(* IEC 61131-3 sources: plc-st-coding-agent/progress/evidence/f14_v14_remaining_20261113/jobs/codex_deepseek-v4pro (part 3) *)

(* ---- public-hard-05.candidate_02.st ---- *)
(* ENGINEERING_CONTRACT
   Manual axis output: ON while its button=1, opposite command inactive, and its limit=0; OFF on release/limit (PUB001).
   Manual grip/release: ON while button=1, opposite inactive, and its limit=0; OFF on release/limit (PUB001).
   Single-step: Start edge activates next index 0..7/wraps; output held until switch; next Start advances (PUB002-PUB003).
   Single-cycle: Start edge runs 0..7; holds each output until completion; stops after left; next Start restarts (PUB004).
   Continuous: Start edge runs 0..7 and loops after left while mode selected (PUB005).
   Emergency: EmergencyStop=FALSE overrides all outputs and freezes start/progression; state is retained (PUB006).
   Index completion: 0/4 DownLimit, 1 GripLimit, 2/6 UpLimit, 3 RightLimit, 5 ReleaseLimit, 7 LeftLimit.
   Same-scan priority: E-stop highest; sequential completion advances the step before output evaluation, so the next action can start on the completed action's scan.
   Unspecified: post-E-stop resumption uses retained state; mode changes outside a mode retain sequence state.
*)
(* CONTRACT_RULES [] *)

FUNCTION_BLOCK MechanicalArmControl
VAR_INPUT
    ManualMode : BOOL;
    SingleStepMode : BOOL;
    SingleCycleMode : BOOL;
    ContinuousMode : BOOL;
    EmergencyStop : BOOL;
    Start : BOOL;
    DownButton : BOOL;
    UpButton : BOOL;
    LeftButton : BOOL;
    RightButton : BOOL;
    GripButton : BOOL;
    ReleaseButton : BOOL;
    DownLimitSwitch : BOOL;
    UpLimitSwitch : BOOL;
    LeftLimitSwitch : BOOL;
    RightLimitSwitch : BOOL;
    GripLimitSwitch : BOOL;
    ReleaseLimitSwitch : BOOL;
END_VAR
VAR_OUTPUT
    MoveDown : BOOL;
    MoveUp : BOOL;
    MoveLeft : BOOL;
    MoveRight : BOOL;
    ActivateGrip : BOOL;
    ActivateRelease : BOOL;
END_VAR
VAR
    tmp_startEdge : R_TRIG;
    tmp_autoMode : BOOL;
    tmp_autoActive : BOOL := FALSE;
    tmp_currentStep : INT := 0;
    tmp_singleNextStep : INT := 0;
    tmp_targetReached : BOOL;
    tmp_prevSelectedModeKey : INT := -1;
    tmp_selectedModeKey : INT;

    tmp_manualDownReq : BOOL;
    tmp_manualUpReq : BOOL;
    tmp_manualLeftReq : BOOL;
    tmp_manualRightReq : BOOL;
    tmp_manualGripReq : BOOL;
    tmp_manualReleaseReq : BOOL;

    tmp_autoDown : BOOL;
    tmp_autoUp : BOOL;
    tmp_autoLeft : BOOL;
    tmp_autoRight : BOOL;
    tmp_autoGrip : BOOL;
    tmp_autoRelease : BOOL;

    tmp_down : BOOL;
    tmp_up : BOOL;
    tmp_left : BOOL;
    tmp_right : BOOL;
    tmp_grip : BOOL;
    tmp_release : BOOL;
END_VAR

tmp_startEdge(CLK := Start);

tmp_manualDownReq := ManualMode AND DownButton AND NOT DownLimitSwitch;
tmp_manualUpReq := ManualMode AND UpButton AND NOT UpLimitSwitch;
tmp_manualLeftReq := ManualMode AND LeftButton AND NOT LeftLimitSwitch;
tmp_manualRightReq := ManualMode AND RightButton AND NOT RightLimitSwitch;
tmp_manualGripReq := ManualMode AND GripButton AND NOT GripLimitSwitch;
tmp_manualReleaseReq := ManualMode AND ReleaseButton AND NOT ReleaseLimitSwitch;

tmp_autoMode := SingleStepMode OR SingleCycleMode OR ContinuousMode;

tmp_selectedModeKey := 0;
IF SingleStepMode THEN
    tmp_selectedModeKey := 1;
ELSIF SingleCycleMode THEN
    tmp_selectedModeKey := 2;
ELSIF ContinuousMode THEN
    tmp_selectedModeKey := 3;
END_IF;

IF tmp_selectedModeKey <> tmp_prevSelectedModeKey THEN
    tmp_autoActive := FALSE;
    tmp_currentStep := 0;
END_IF;
tmp_prevSelectedModeKey := tmp_selectedModeKey;

IF EmergencyStop AND tmp_startEdge.Q THEN
    IF SingleStepMode THEN
        IF NOT tmp_autoActive THEN
            tmp_currentStep := tmp_singleNextStep;
            tmp_singleNextStep := (tmp_singleNextStep + 1) MOD 8;
            tmp_autoActive := TRUE;
        END_IF;
    ELSIF SingleCycleMode THEN
        IF NOT tmp_autoActive THEN
            tmp_currentStep := 0;
            tmp_autoActive := TRUE;
        END_IF;
    ELSIF ContinuousMode THEN
        IF NOT tmp_autoActive THEN
            tmp_currentStep := 0;
            tmp_autoActive := TRUE;
        END_IF;
    END_IF;
END_IF;

CASE tmp_currentStep OF
    0, 4:
        tmp_targetReached := DownLimitSwitch;
    1:
        tmp_targetReached := GripLimitSwitch;
    2, 6:
        tmp_targetReached := UpLimitSwitch;
    3:
        tmp_targetReached := RightLimitSwitch;
    5:
        tmp_targetReached := ReleaseLimitSwitch;
    7:
        tmp_targetReached := LeftLimitSwitch;
ELSE
    tmp_targetReached := FALSE;
END_CASE;

IF EmergencyStop AND tmp_autoMode AND tmp_autoActive AND tmp_targetReached THEN
    IF SingleStepMode THEN
        tmp_autoActive := FALSE;
    ELSIF SingleCycleMode THEN
        IF tmp_currentStep >= 7 THEN
            tmp_autoActive := FALSE;
            tmp_currentStep := 0;
        ELSE
            tmp_currentStep := tmp_currentStep + 1;
        END_IF;
    ELSIF ContinuousMode THEN
        IF tmp_currentStep >= 7 THEN
            tmp_currentStep := 0;
        ELSE
            tmp_currentStep := tmp_currentStep + 1;
        END_IF;
    END_IF;
END_IF;

tmp_autoDown := tmp_autoMode AND tmp_autoActive AND ((tmp_currentStep = 0) OR (tmp_currentStep = 4)) AND NOT DownLimitSwitch;
tmp_autoGrip := tmp_autoMode AND tmp_autoActive AND (tmp_currentStep = 1) AND NOT GripLimitSwitch;
tmp_autoUp := tmp_autoMode AND tmp_autoActive AND ((tmp_currentStep = 2) OR (tmp_currentStep = 6)) AND NOT UpLimitSwitch;
tmp_autoRight := tmp_autoMode AND tmp_autoActive AND (tmp_currentStep = 3) AND NOT RightLimitSwitch;
tmp_autoRelease := tmp_autoMode AND tmp_autoActive AND (tmp_currentStep = 5) AND NOT ReleaseLimitSwitch;
tmp_autoLeft := tmp_autoMode AND tmp_autoActive AND (tmp_currentStep = 7) AND NOT LeftLimitSwitch;

tmp_down := tmp_manualDownReq OR tmp_autoDown;
tmp_up := tmp_manualUpReq OR tmp_autoUp;
tmp_left := tmp_manualLeftReq OR tmp_autoLeft;
tmp_right := tmp_manualRightReq OR tmp_autoRight;
tmp_grip := tmp_manualGripReq OR tmp_autoGrip;
tmp_release := tmp_manualReleaseReq OR tmp_autoRelease;

MoveDown := tmp_down AND NOT tmp_up AND EmergencyStop;
MoveUp := tmp_up AND NOT tmp_down AND EmergencyStop;
MoveLeft := tmp_left AND NOT tmp_right AND EmergencyStop;
MoveRight := tmp_right AND NOT tmp_left AND EmergencyStop;
ActivateGrip := tmp_grip AND NOT tmp_release AND EmergencyStop;
ActivateRelease := tmp_release AND NOT tmp_grip AND EmergencyStop;

END_FUNCTION_BLOCK

(* ---- public-hard-05.patch_base_02.st ---- *)
(* ENGINEERING_CONTRACT
   Manual axis output: ON while its button=1, opposite command inactive, and its limit=0; OFF on release/limit (PUB001).
   Manual grip/release: ON while button=1, opposite inactive, and its limit=0; OFF on release/limit (PUB001).
   Single-step: Start edge activates next index 0..7/wraps; output held until switch; next Start advances (PUB002-PUB003).
   Single-cycle: Start edge runs 0..7; holds each output until completion; stops after left; next Start restarts (PUB004).
   Continuous: Start edge runs 0..7 and loops after left while mode selected (PUB005).
   Emergency: EmergencyStop=FALSE overrides all outputs and freezes start/progression; state is retained (PUB006).
   Index completion: 0/4 DownLimit, 1 GripLimit, 2/6 UpLimit, 3 RightLimit, 5 ReleaseLimit, 7 LeftLimit.
   Same-scan priority: E-stop highest; a feedback-completed action cannot energize on its completion scan; next action starts next scan.
   Unspecified: post-E-stop resumption uses retained state; mode changes outside a mode retain sequence state.
*)
(* CONTRACT_RULES [] *)

FUNCTION_BLOCK MechanicalArmControl
VAR_INPUT
    ManualMode : BOOL;
    SingleStepMode : BOOL;
    SingleCycleMode : BOOL;
    ContinuousMode : BOOL;
    EmergencyStop : BOOL;
    Start : BOOL;
    DownButton : BOOL;
    UpButton : BOOL;
    LeftButton : BOOL;
    RightButton : BOOL;
    GripButton : BOOL;
    ReleaseButton : BOOL;
    DownLimitSwitch : BOOL;
    UpLimitSwitch : BOOL;
    LeftLimitSwitch : BOOL;
    RightLimitSwitch : BOOL;
    GripLimitSwitch : BOOL;
    ReleaseLimitSwitch : BOOL;
END_VAR
VAR_OUTPUT
    MoveDown : BOOL;
    MoveUp : BOOL;
    MoveLeft : BOOL;
    MoveRight : BOOL;
    ActivateGrip : BOOL;
    ActivateRelease : BOOL;
END_VAR
VAR
    tmp_startEdge : R_TRIG;
    tmp_autoMode : BOOL;
    tmp_autoActive : BOOL := FALSE;
    tmp_currentStep : INT := 0;
    tmp_singleNextStep : INT := 0;
    tmp_targetReached : BOOL;

    tmp_manualDownReq : BOOL;
    tmp_manualUpReq : BOOL;
    tmp_manualLeftReq : BOOL;
    tmp_manualRightReq : BOOL;
    tmp_manualGripReq : BOOL;
    tmp_manualReleaseReq : BOOL;

    tmp_autoDown : BOOL;
    tmp_autoUp : BOOL;
    tmp_autoLeft : BOOL;
    tmp_autoRight : BOOL;
    tmp_autoGrip : BOOL;
    tmp_autoRelease : BOOL;

    tmp_down : BOOL;
    tmp_up : BOOL;
    tmp_left : BOOL;
    tmp_right : BOOL;
    tmp_grip : BOOL;
    tmp_release : BOOL;
END_VAR

tmp_startEdge(CLK := Start);

tmp_manualDownReq := ManualMode AND DownButton AND NOT DownLimitSwitch;
tmp_manualUpReq := ManualMode AND UpButton AND NOT UpLimitSwitch;
tmp_manualLeftReq := ManualMode AND LeftButton AND NOT LeftLimitSwitch;
tmp_manualRightReq := ManualMode AND RightButton AND NOT RightLimitSwitch;
tmp_manualGripReq := ManualMode AND GripButton AND NOT GripLimitSwitch;
tmp_manualReleaseReq := ManualMode AND ReleaseButton AND NOT ReleaseLimitSwitch;

tmp_autoMode := SingleStepMode OR SingleCycleMode OR ContinuousMode;

IF EmergencyStop AND tmp_startEdge.Q THEN
    IF SingleStepMode THEN
        IF NOT tmp_autoActive THEN
            tmp_currentStep := tmp_singleNextStep;
            tmp_singleNextStep := (tmp_singleNextStep + 1) MOD 8;
            tmp_autoActive := TRUE;
        END_IF;
    ELSIF SingleCycleMode THEN
        IF NOT tmp_autoActive THEN
            tmp_currentStep := 0;
            tmp_autoActive := TRUE;
        END_IF;
    ELSIF ContinuousMode THEN
        IF NOT tmp_autoActive THEN
            tmp_currentStep := 0;
            tmp_autoActive := TRUE;
        END_IF;
    END_IF;
END_IF;

CASE tmp_currentStep OF
    0, 4:
        tmp_targetReached := DownLimitSwitch;
    1:
        tmp_targetReached := GripLimitSwitch;
    2, 6:
        tmp_targetReached := UpLimitSwitch;
    3:
        tmp_targetReached := RightLimitSwitch;
    5:
        tmp_targetReached := ReleaseLimitSwitch;
    7:
        tmp_targetReached := LeftLimitSwitch;
ELSE
    tmp_targetReached := FALSE;
END_CASE;

tmp_autoDown := tmp_autoMode AND tmp_autoActive AND ((tmp_currentStep = 0) OR (tmp_currentStep = 4)) AND NOT DownLimitSwitch;
tmp_autoGrip := tmp_autoMode AND tmp_autoActive AND (tmp_currentStep = 1) AND NOT GripLimitSwitch;
tmp_autoUp := tmp_autoMode AND tmp_autoActive AND ((tmp_currentStep = 2) OR (tmp_currentStep = 6)) AND NOT UpLimitSwitch;
tmp_autoRight := tmp_autoMode AND tmp_autoActive AND (tmp_currentStep = 3) AND NOT RightLimitSwitch;
tmp_autoRelease := tmp_autoMode AND tmp_autoActive AND (tmp_currentStep = 5) AND NOT ReleaseLimitSwitch;
tmp_autoLeft := tmp_autoMode AND tmp_autoActive AND (tmp_currentStep = 7) AND NOT LeftLimitSwitch;

tmp_down := tmp_manualDownReq OR tmp_autoDown;
tmp_up := tmp_manualUpReq OR tmp_autoUp;
tmp_left := tmp_manualLeftReq OR tmp_autoLeft;
tmp_right := tmp_manualRightReq OR tmp_autoRight;
tmp_grip := tmp_manualGripReq OR tmp_autoGrip;
tmp_release := tmp_manualReleaseReq OR tmp_autoRelease;

MoveDown := tmp_down AND NOT tmp_up AND EmergencyStop;
MoveUp := tmp_up AND NOT tmp_down AND EmergencyStop;
MoveLeft := tmp_left AND NOT tmp_right AND EmergencyStop;
MoveRight := tmp_right AND NOT tmp_left AND EmergencyStop;
ActivateGrip := tmp_grip AND NOT tmp_release AND EmergencyStop;
ActivateRelease := tmp_release AND NOT tmp_grip AND EmergencyStop;

IF EmergencyStop AND tmp_autoMode AND tmp_autoActive AND tmp_targetReached THEN
    IF SingleStepMode THEN
        tmp_autoActive := FALSE;
    ELSIF SingleCycleMode THEN
        IF tmp_currentStep >= 7 THEN
            tmp_autoActive := FALSE;
            tmp_currentStep := 0;
        ELSE
            tmp_currentStep := tmp_currentStep + 1;
        END_IF;
    ELSIF ContinuousMode THEN
        IF tmp_currentStep >= 7 THEN
            tmp_currentStep := 0;
        ELSE
            tmp_currentStep := tmp_currentStep + 1;
        END_IF;
    END_IF;
END_IF;

END_FUNCTION_BLOCK

(* ---- public-hard-05.raw_candidate_01.st ---- *)
(* ENGINEERING_CONTRACT
   Manual axis output: ON while its button=1, opposite command inactive, and its limit=0; OFF on release/limit (PUB001).
   Manual grip/release: ON while button=1, opposite inactive, and its limit=0; OFF on release/limit (PUB001).
   Single-step: Start edge activates next index 0..7/wraps; output held until switch; next Start advances (PUB002-PUB003).
   Single-cycle: Start edge runs 0..7; holds each output until completion; stops after left; next Start restarts (PUB004).
   Continuous: Start edge runs 0..7 and loops after left while mode selected (PUB005).
   Emergency: EmergencyStop=FALSE overrides all outputs and freezes start/progression; state is retained (PUB006).
   Index completion: 0/4 DownLimit, 1 GripLimit, 2/6 UpLimit, 3 RightLimit, 5 ReleaseLimit, 7 LeftLimit.
   Same-scan priority: E-stop highest; a feedback-completed action cannot energize on its completion scan; next action starts next scan.
   Unspecified: post-E-stop resumption uses retained state; mode changes outside a mode retain sequence state.
*)
(* CONTRACT_RULES [] *)

FUNCTION_BLOCK MechanicalArmControl
VAR_INPUT
    ManualMode : BOOL;
    SingleStepMode : BOOL;
    SingleCycleMode : BOOL;
    ContinuousMode : BOOL;
    EmergencyStop : BOOL;
    Start : BOOL;
    DownButton : BOOL;
    UpButton : BOOL;
    LeftButton : BOOL;
    RightButton : BOOL;
    GripButton : BOOL;
    ReleaseButton : BOOL;
    DownLimitSwitch : BOOL;
    UpLimitSwitch : BOOL;
    LeftLimitSwitch : BOOL;
    RightLimitSwitch : BOOL;
    GripLimitSwitch : BOOL;
    ReleaseLimitSwitch : BOOL;
END_VAR
VAR_OUTPUT
    MoveDown : BOOL;
    MoveUp : BOOL;
    MoveLeft : BOOL;
    MoveRight : BOOL;
    ActivateGrip : BOOL;
    ActivateRelease : BOOL;
END_VAR
VAR
    tmp_startEdge : R_TRIG;
    tmp_autoMode : BOOL;
    tmp_autoActive : BOOL := FALSE;
    tmp_currentStep : INT := 0;
    tmp_singleNextStep : INT := 0;
    tmp_targetReached : BOOL;

    tmp_manualDownReq : BOOL;
    tmp_manualUpReq : BOOL;
    tmp_manualLeftReq : BOOL;
    tmp_manualRightReq : BOOL;
    tmp_manualGripReq : BOOL;
    tmp_manualReleaseReq : BOOL;

    tmp_autoDown : BOOL;
    tmp_autoUp : BOOL;
    tmp_autoLeft : BOOL;
    tmp_autoRight : BOOL;
    tmp_autoGrip : BOOL;
    tmp_autoRelease : BOOL;

    tmp_down : BOOL;
    tmp_up : BOOL;
    tmp_left : BOOL;
    tmp_right : BOOL;
    tmp_grip : BOOL;
    tmp_release : BOOL;
END_VAR

tmp_startEdge(CLK := Start);

tmp_manualDownReq := ManualMode AND DownButton AND NOT DownLimitSwitch;
tmp_manualUpReq := ManualMode AND UpButton AND NOT UpLimitSwitch;
tmp_manualLeftReq := ManualMode AND LeftButton AND NOT LeftLimitSwitch;
tmp_manualRightReq := ManualMode AND RightButton AND NOT RightLimitSwitch;
tmp_manualGripReq := ManualMode AND GripButton AND NOT GripLimitSwitch;
tmp_manualReleaseReq := ManualMode AND ReleaseButton AND NOT ReleaseLimitSwitch;

tmp_autoMode := SingleStepMode OR SingleCycleMode OR ContinuousMode;

IF EmergencyStop AND tmp_startEdge.Q THEN
    IF SingleStepMode THEN
        IF NOT tmp_autoActive THEN
            tmp_currentStep := tmp_singleNextStep;
            tmp_singleNextStep := (tmp_singleNextStep + 1) MOD 8;
            tmp_autoActive := TRUE;
        END_IF;
    ELSIF SingleCycleMode THEN
        IF NOT tmp_autoActive THEN
            tmp_currentStep := 0;
            tmp_autoActive := TRUE;
        END_IF;
    ELSIF ContinuousMode THEN
        IF NOT tmp_autoActive THEN
            tmp_currentStep := 0;
            tmp_autoActive := TRUE;
        END_IF;
    END_IF;
END_IF;

CASE tmp_currentStep OF
    0, 4:
        tmp_targetReached := DownLimitSwitch;
    1:
        tmp_targetReached := GripLimitSwitch;
    2, 6:
        tmp_targetReached := UpLimitSwitch;
    3:
        tmp_targetReached := RightLimitSwitch;
    5:
        tmp_targetReached := ReleaseLimitSwitch;
    7:
        tmp_targetReached := LeftLimitSwitch;
ELSE
    tmp_targetReached := FALSE;
END_CASE;

tmp_autoDown := tmp_autoMode AND tmp_autoActive AND ((tmp_currentStep = 0) OR (tmp_currentStep = 4)) AND NOT DownLimitSwitch;
tmp_autoGrip := tmp_autoMode AND tmp_autoActive AND (tmp_currentStep = 1) AND NOT GripLimitSwitch;
tmp_autoUp := tmp_autoMode AND tmp_autoActive AND ((tmp_currentStep = 2) OR (tmp_currentStep = 6)) AND NOT UpLimitSwitch;
tmp_autoRight := tmp_autoMode AND tmp_autoActive AND (tmp_currentStep = 3) AND NOT RightLimitSwitch;
tmp_autoRelease := tmp_autoMode AND tmp_autoActive AND (tmp_currentStep = 5) AND NOT ReleaseLimitSwitch;
tmp_autoLeft := tmp_autoMode AND tmp_autoActive AND (tmp_currentStep = 7) AND NOT LeftLimitSwitch;

tmp_down := tmp_manualDownReq OR tmp_autoDown;
tmp_up := tmp_manualUpReq OR tmp_autoUp;
tmp_left := tmp_manualLeftReq OR tmp_autoLeft;
tmp_right := tmp_manualRightReq OR tmp_autoRight;
tmp_grip := tmp_manualGripReq OR tmp_autoGrip;
tmp_release := tmp_manualReleaseReq OR tmp_autoRelease;

MoveDown := tmp_down AND NOT tmp_up AND EmergencyStop;
MoveUp := tmp_up AND NOT tmp_down AND EmergencyStop;
MoveLeft := tmp_left AND NOT tmp_right AND EmergencyStop;
MoveRight := tmp_right AND NOT tmp_left AND EmergencyStop;
ActivateGrip := tmp_grip AND NOT tmp_release AND EmergencyStop;
ActivateRelease := tmp_release AND NOT tmp_grip AND EmergencyStop;

IF EmergencyStop AND tmp_autoMode AND tmp_autoActive AND tmp_targetReached THEN
    IF SingleStepMode THEN
        tmp_autoActive := FALSE;
    ELSIF SingleCycleMode THEN
        IF tmp_currentStep >= 7 THEN
            tmp_autoActive := FALSE;
            tmp_currentStep := 0;
        ELSE
            tmp_currentStep := tmp_currentStep + 1;
        END_IF;
    ELSIF ContinuousMode THEN
        IF tmp_currentStep >= 7 THEN
            tmp_currentStep := 0;
        ELSE
            tmp_currentStep := tmp_currentStep + 1;
        END_IF;
    END_IF;
END_IF;

END_FUNCTION_BLOCK

(* ---- public-hard-05.raw_candidate_02.st ---- *)
(* ENGINEERING_CONTRACT
   Manual axis output: ON while its button=1, opposite command inactive, and its limit=0; OFF on release/limit (PUB001).
   Manual grip/release: ON while button=1, opposite inactive, and its limit=0; OFF on release/limit (PUB001).
   Single-step: Start edge activates next index 0..7/wraps; output held until switch; next Start advances (PUB002-PUB003).
   Single-cycle: Start edge runs 0..7; holds each output until completion; stops after left; next Start restarts (PUB004).
   Continuous: Start edge runs 0..7 and loops after left while mode selected (PUB005).
   Emergency: EmergencyStop=FALSE overrides all outputs and freezes start/progression; state is retained (PUB006).
   Index completion: 0/4 DownLimit, 1 GripLimit, 2/6 UpLimit, 3 RightLimit, 5 ReleaseLimit, 7 LeftLimit.
   Same-scan priority: E-stop highest; sequential completion advances the step before output evaluation, so the next action can start on the completed action's scan.
   Unspecified: post-E-stop resumption uses retained state; mode changes outside a mode retain sequence state.
*)
(* CONTRACT_RULES [] *)

FUNCTION_BLOCK MechanicalArmControl
VAR_INPUT
    ManualMode : BOOL;
    SingleStepMode : BOOL;
    SingleCycleMode : BOOL;
    ContinuousMode : BOOL;
    EmergencyStop : BOOL;
    Start : BOOL;
    DownButton : BOOL;
    UpButton : BOOL;
    LeftButton : BOOL;
    RightButton : BOOL;
    GripButton : BOOL;
    ReleaseButton : BOOL;
    DownLimitSwitch : BOOL;
    UpLimitSwitch : BOOL;
    LeftLimitSwitch : BOOL;
    RightLimitSwitch : BOOL;
    GripLimitSwitch : BOOL;
    ReleaseLimitSwitch : BOOL;
END_VAR
VAR_OUTPUT
    MoveDown : BOOL;
    MoveUp : BOOL;
    MoveLeft : BOOL;
    MoveRight : BOOL;
    ActivateGrip : BOOL;
    ActivateRelease : BOOL;
END_VAR
VAR
    tmp_startEdge : R_TRIG;
    tmp_autoMode : BOOL;
    tmp_autoActive : BOOL := FALSE;
    tmp_currentStep : INT := 0;
    tmp_singleNextStep : INT := 0;
    tmp_targetReached : BOOL;
    tmp_prevSelectedModeKey : INT := -1;
    tmp_selectedModeKey : INT;

    tmp_manualDownReq : BOOL;
    tmp_manualUpReq : BOOL;
    tmp_manualLeftReq : BOOL;
    tmp_manualRightReq : BOOL;
    tmp_manualGripReq : BOOL;
    tmp_manualReleaseReq : BOOL;

    tmp_autoDown : BOOL;
    tmp_autoUp : BOOL;
    tmp_autoLeft : BOOL;
    tmp_autoRight : BOOL;
    tmp_autoGrip : BOOL;
    tmp_autoRelease : BOOL;

    tmp_down : BOOL;
    tmp_up : BOOL;
    tmp_left : BOOL;
    tmp_right : BOOL;
    tmp_grip : BOOL;
    tmp_release : BOOL;
END_VAR

tmp_startEdge(CLK := Start);

tmp_manualDownReq := ManualMode AND DownButton AND NOT DownLimitSwitch;
tmp_manualUpReq := ManualMode AND UpButton AND NOT UpLimitSwitch;
tmp_manualLeftReq := ManualMode AND LeftButton AND NOT LeftLimitSwitch;
tmp_manualRightReq := ManualMode AND RightButton AND NOT RightLimitSwitch;
tmp_manualGripReq := ManualMode AND GripButton AND NOT GripLimitSwitch;
tmp_manualReleaseReq := ManualMode AND ReleaseButton AND NOT ReleaseLimitSwitch;

tmp_autoMode := SingleStepMode OR SingleCycleMode OR ContinuousMode;

tmp_selectedModeKey := 0;
IF SingleStepMode THEN
    tmp_selectedModeKey := 1;
ELSIF SingleCycleMode THEN
    tmp_selectedModeKey := 2;
ELSIF ContinuousMode THEN
    tmp_selectedModeKey := 3;
END_IF;

IF tmp_selectedModeKey <> tmp_prevSelectedModeKey THEN
    tmp_autoActive := FALSE;
    tmp_currentStep := 0;
END_IF;
tmp_prevSelectedModeKey := tmp_selectedModeKey;

IF EmergencyStop AND tmp_startEdge.Q THEN
    IF SingleStepMode THEN
        IF NOT tmp_autoActive THEN
            tmp_currentStep := tmp_singleNextStep;
            tmp_singleNextStep := (tmp_singleNextStep + 1) MOD 8;
            tmp_autoActive := TRUE;
        END_IF;
    ELSIF SingleCycleMode THEN
        IF NOT tmp_autoActive THEN
            tmp_currentStep := 0;
            tmp_autoActive := TRUE;
        END_IF;
    ELSIF ContinuousMode THEN
        IF NOT tmp_autoActive THEN
            tmp_currentStep := 0;
            tmp_autoActive := TRUE;
        END_IF;
    END_IF;
END_IF;

CASE tmp_currentStep OF
    0, 4:
        tmp_targetReached := DownLimitSwitch;
    1:
        tmp_targetReached := GripLimitSwitch;
    2, 6:
        tmp_targetReached := UpLimitSwitch;
    3:
        tmp_targetReached := RightLimitSwitch;
    5:
        tmp_targetReached := ReleaseLimitSwitch;
    7:
        tmp_targetReached := LeftLimitSwitch;
ELSE
    tmp_targetReached := FALSE;
END_CASE;

IF EmergencyStop AND tmp_autoMode AND tmp_autoActive AND tmp_targetReached THEN
    IF SingleStepMode THEN
        tmp_autoActive := FALSE;
    ELSIF SingleCycleMode THEN
        IF tmp_currentStep >= 7 THEN
            tmp_autoActive := FALSE;
            tmp_currentStep := 0;
        ELSE
            tmp_currentStep := tmp_currentStep + 1;
        END_IF;
    ELSIF ContinuousMode THEN
        IF tmp_currentStep >= 7 THEN
            tmp_currentStep := 0;
        ELSE
            tmp_currentStep := tmp_currentStep + 1;
        END_IF;
    END_IF;
END_IF;

tmp_autoDown := tmp_autoMode AND tmp_autoActive AND ((tmp_currentStep = 0) OR (tmp_currentStep = 4)) AND NOT DownLimitSwitch;
tmp_autoGrip := tmp_autoMode AND tmp_autoActive AND (tmp_currentStep = 1) AND NOT GripLimitSwitch;
tmp_autoUp := tmp_autoMode AND tmp_autoActive AND ((tmp_currentStep = 2) OR (tmp_currentStep = 6)) AND NOT UpLimitSwitch;
tmp_autoRight := tmp_autoMode AND tmp_autoActive AND (tmp_currentStep = 3) AND NOT RightLimitSwitch;
tmp_autoRelease := tmp_autoMode AND tmp_autoActive AND (tmp_currentStep = 5) AND NOT ReleaseLimitSwitch;
tmp_autoLeft := tmp_autoMode AND tmp_autoActive AND (tmp_currentStep = 7) AND NOT LeftLimitSwitch;

tmp_down := tmp_manualDownReq OR tmp_autoDown;
tmp_up := tmp_manualUpReq OR tmp_autoUp;
tmp_left := tmp_manualLeftReq OR tmp_autoLeft;
tmp_right := tmp_manualRightReq OR tmp_autoRight;
tmp_grip := tmp_manualGripReq OR tmp_autoGrip;
tmp_release := tmp_manualReleaseReq OR tmp_autoRelease;

MoveDown := tmp_down AND NOT tmp_up AND EmergencyStop;
MoveUp := tmp_up AND NOT tmp_down AND EmergencyStop;
MoveLeft := tmp_left AND NOT tmp_right AND EmergencyStop;
MoveRight := tmp_right AND NOT tmp_left AND EmergencyStop;
ActivateGrip := tmp_grip AND NOT tmp_release AND EmergencyStop;
ActivateRelease := tmp_release AND NOT tmp_grip AND EmergencyStop;

END_FUNCTION_BLOCK

(* ---- public-hard-06.candidate_01.st ---- *)
(* ENGINEERING_CONTRACT
- MotorForward/MotorReverse: manual direct from buttons, both inhibited when both are requested or Mode=1; automatic uses forward motion states only (PUB001, PUB002).
- Automatic motion: enabled by feed/cleaning/weighing/firing completion and held until the destination sensor is active; same-scan arrival has priority over completion (PUB003-PUB008).
- kick: set when weighing completes with weight<100.0 or weight>200.0; held while rejected until SensorWeight clears or Mode=0 (PUB009).
- firingTemp: updated only on a qualified weighing, REAL degrees, linear 100..200 -> 500..550; held through firing/output until unqualified, next feed, or Mode=0 (PUB009, PUB010).
- CompletionLight: active while SensorOutput in automatic output state; cleared when the product is removed or Mode=0 (PUB008).
- Weight boundary test is inclusive: qualified is 100.0 <= weight <= 200.0 (PUB009).
*)
(* CONTRACT_RULES [] *)

TYPE E_ProductionState :
(
    ST_IDLE := 0,
    ST_MOVE_TO_WASH := 1,
    ST_AT_WASH := 2,
    ST_MOVE_TO_WEIGHT := 3,
    ST_AT_WEIGHT := 4,
    ST_MOVE_TO_FIRING := 5,
    ST_AT_FIRING := 6,
    ST_MOVE_TO_OUTPUT := 7,
    ST_AT_OUTPUT := 8,
    ST_REJECTED := 9
);
END_TYPE;

FUNCTION_BLOCK ProductionControl
VAR_INPUT
    Mode : BOOL;
    ForwardButton : BOOL;
    ReverseButton : BOOL;
    SensorFeed : BOOL;
    SensorWash : BOOL;
    SensorWeight : BOOL;
    SensorFiring : BOOL;
    SensorOutput : BOOL;
    washComplete : BOOL;
    weightComplete : BOOL;
    weight : REAL;
    firingComplete : BOOL;
END_VAR
VAR_OUTPUT
    MotorForward : BOOL;
    MotorReverse : BOOL;
    kick : BOOL;
    CompletionLight : BOOL;
    firingTemp : REAL;
END_VAR
VAR
    tmp_LocalState : E_ProductionState := ST_IDLE;
    tmp_Qualified : BOOL;
    tmp_TempLatched : REAL := 0.0;
END_VAR

IF NOT Mode THEN
    MotorForward := ForwardButton AND NOT ReverseButton;
    MotorReverse := ReverseButton AND NOT ForwardButton;
    kick := FALSE;
    CompletionLight := FALSE;
    tmp_TempLatched := 0.0;
    firingTemp := 0.0;
ELSE
    MotorReverse := FALSE;

    IF tmp_LocalState = ST_IDLE THEN
        tmp_TempLatched := 0.0;
        IF SensorFeed THEN
            tmp_LocalState := ST_MOVE_TO_WASH;
        END_IF;
    ELSIF tmp_LocalState = ST_MOVE_TO_WASH THEN
        IF SensorWash THEN
            tmp_LocalState := ST_AT_WASH;
        END_IF;
    ELSIF tmp_LocalState = ST_AT_WASH THEN
        IF SensorWeight THEN
            tmp_LocalState := ST_AT_WEIGHT;
        ELSIF washComplete THEN
            tmp_LocalState := ST_MOVE_TO_WEIGHT;
        END_IF;
    ELSIF tmp_LocalState = ST_MOVE_TO_WEIGHT THEN
        IF SensorWeight THEN
            tmp_LocalState := ST_AT_WEIGHT;
        END_IF;
    ELSIF tmp_LocalState = ST_AT_WEIGHT THEN
        IF SensorFiring THEN
            tmp_LocalState := ST_AT_FIRING;
        ELSIF weightComplete THEN
            tmp_Qualified := (weight >= 100.0) AND (weight <= 200.0);
            IF tmp_Qualified THEN
                tmp_TempLatched := 500.0 + ((weight - 100.0) * 50.0) / 100.0;
                tmp_LocalState := ST_MOVE_TO_FIRING;
            ELSE
                tmp_TempLatched := 0.0;
                tmp_LocalState := ST_REJECTED;
            END_IF;
        END_IF;
    ELSIF tmp_LocalState = ST_REJECTED THEN
        IF NOT SensorWeight THEN
            tmp_TempLatched := 0.0;
            tmp_LocalState := ST_IDLE;
        END_IF;
    ELSIF tmp_LocalState = ST_MOVE_TO_FIRING THEN
        IF SensorFiring THEN
            tmp_LocalState := ST_AT_FIRING;
        END_IF;
    ELSIF tmp_LocalState = ST_AT_FIRING THEN
        IF SensorOutput THEN
            tmp_LocalState := ST_AT_OUTPUT;
        ELSIF firingComplete THEN
            tmp_LocalState := ST_MOVE_TO_OUTPUT;
        END_IF;
    ELSIF tmp_LocalState = ST_MOVE_TO_OUTPUT THEN
        IF SensorOutput THEN
            tmp_LocalState := ST_AT_OUTPUT;
        END_IF;
    ELSIF tmp_LocalState = ST_AT_OUTPUT THEN
        IF NOT SensorOutput THEN
            tmp_TempLatched := 0.0;
            tmp_LocalState := ST_IDLE;
        END_IF;
    END_IF;

    CASE tmp_LocalState OF
        ST_MOVE_TO_WASH,
        ST_MOVE_TO_WEIGHT,
        ST_MOVE_TO_FIRING,
        ST_MOVE_TO_OUTPUT:
            MotorForward := TRUE;
    ELSE
            MotorForward := FALSE;
    END_CASE;

    kick := (tmp_LocalState = ST_REJECTED);
    CompletionLight := (tmp_LocalState = ST_AT_OUTPUT) AND SensorOutput;
    firingTemp := tmp_TempLatched;
END_IF;

(* ---- public-hard-06.candidate_02.st ---- *)
(* ENGINEERING_CONTRACT
- MotorForward/MotorReverse: manual direct from buttons, both inhibited when both are requested or Mode=1; automatic uses forward motion states only (PUB001, PUB002).
- Automatic motion: enabled by feed/cleaning/weighing/firing completion and held until the destination sensor is active; same-scan arrival has priority over completion (PUB003-PUB008).
- kick: set when weighing completes with weight<100.0 or weight>200.0; held while rejected until SensorWeight clears or Mode=0 (PUB009).
- firingTemp: updated only on a qualified weighing, REAL degrees, linear 100..200 -> 500..550; held through firing/output until unqualified, next feed, or Mode=0 (PUB009, PUB010).
- CompletionLight: active while SensorOutput in automatic output state; cleared when the product is removed or Mode=0 (PUB008).
- Weight boundary test is inclusive: qualified is 100.0 <= weight <= 200.0 (PUB009).
*)
(* CONTRACT_RULES [] *)

TYPE E_ProductionState :
(
    ST_IDLE := 0,
    ST_MOVE_TO_WASH := 1,
    ST_AT_WASH := 2,
    ST_MOVE_TO_WEIGHT := 3,
    ST_AT_WEIGHT := 4,
    ST_MOVE_TO_FIRING := 5,
    ST_AT_FIRING := 6,
    ST_MOVE_TO_OUTPUT := 7,
    ST_AT_OUTPUT := 8,
    ST_REJECTED := 9
);
END_TYPE;

FUNCTION_BLOCK ProductionControl
VAR_INPUT
    Mode : BOOL;
    ForwardButton : BOOL;
    ReverseButton : BOOL;
    SensorFeed : BOOL;
    SensorWash : BOOL;
    SensorWeight : BOOL;
    SensorFiring : BOOL;
    SensorOutput : BOOL;
    washComplete : BOOL;
    weightComplete : BOOL;
    weight : REAL;
    firingComplete : BOOL;
END_VAR
VAR_OUTPUT
    MotorForward : BOOL;
    MotorReverse : BOOL;
    kick : BOOL;
    CompletionLight : BOOL;
    firingTemp : REAL;
END_VAR
VAR
    tmp_LocalState : E_ProductionState := ST_IDLE;
    tmp_Qualified : BOOL;
    tmp_TempLatched : REAL := 0.0;
END_VAR

IF NOT Mode THEN
    MotorForward := ForwardButton AND NOT ReverseButton;
    MotorReverse := ReverseButton AND NOT ForwardButton;
    kick := FALSE;
    CompletionLight := FALSE;
    tmp_TempLatched := 0.0;
    firingTemp := 0.0;
ELSE
    MotorReverse := FALSE;

    IF tmp_LocalState = ST_IDLE THEN
        tmp_TempLatched := 0.0;
        IF SensorFeed THEN
            tmp_LocalState := ST_MOVE_TO_WASH;
        END_IF;
    ELSIF tmp_LocalState = ST_MOVE_TO_WASH THEN
        IF SensorWash THEN
            tmp_LocalState := ST_AT_WASH;
        END_IF;
    ELSIF tmp_LocalState = ST_AT_WASH THEN
        IF SensorWeight THEN
            tmp_LocalState := ST_AT_WEIGHT;
        ELSIF washComplete THEN
            tmp_LocalState := ST_MOVE_TO_WEIGHT;
        END_IF;
    ELSIF tmp_LocalState = ST_MOVE_TO_WEIGHT THEN
        IF SensorWeight THEN
            tmp_LocalState := ST_AT_WEIGHT;
        END_IF;
    ELSIF tmp_LocalState = ST_AT_WEIGHT THEN
        IF SensorFiring THEN
            tmp_LocalState := ST_AT_FIRING;
        ELSIF weightComplete THEN
            tmp_Qualified := (weight >= 100.0) AND (weight <= 200.0);
            IF tmp_Qualified THEN
                tmp_TempLatched := 500.0 + ((weight - 100.0) * 50.0) / 100.0;
                tmp_LocalState := ST_MOVE_TO_FIRING;
            ELSE
                tmp_TempLatched := 0.0;
                tmp_LocalState := ST_REJECTED;
            END_IF;
        END_IF;
    ELSIF tmp_LocalState = ST_REJECTED THEN
        IF NOT SensorWeight THEN
            tmp_TempLatched := 0.0;
            tmp_LocalState := ST_IDLE;
        END_IF;
    ELSIF tmp_LocalState = ST_MOVE_TO_FIRING THEN
        IF SensorFiring THEN
            tmp_LocalState := ST_AT_FIRING;
        END_IF;
    ELSIF tmp_LocalState = ST_AT_FIRING THEN
        IF SensorOutput THEN
            tmp_LocalState := ST_AT_OUTPUT;
        ELSIF firingComplete THEN
            tmp_LocalState := ST_MOVE_TO_OUTPUT;
        END_IF;
    ELSIF tmp_LocalState = ST_MOVE_TO_OUTPUT THEN
        IF SensorOutput THEN
            tmp_LocalState := ST_AT_OUTPUT;
        END_IF;
    ELSIF tmp_LocalState = ST_AT_OUTPUT THEN
        IF NOT SensorOutput THEN
            tmp_TempLatched := 0.0;
            tmp_LocalState := ST_IDLE;
        END_IF;
    END_IF;

    CASE tmp_LocalState OF
        ST_MOVE_TO_WASH,
        ST_MOVE_TO_WEIGHT,
        ST_MOVE_TO_FIRING,
        ST_MOVE_TO_OUTPUT:
            MotorForward := TRUE;
    ELSE
            MotorForward := FALSE;
    END_CASE;

    kick := (tmp_LocalState = ST_REJECTED);
    CompletionLight := (tmp_LocalState = ST_AT_OUTPUT) AND SensorOutput;
    firingTemp := tmp_TempLatched;
END_IF;
END_FUNCTION_BLOCK

(* ---- public-hard-06.candidate_03.st ---- *)
(* ENGINEERING_CONTRACT
- MotorForward/MotorReverse: manual direct from buttons, both inhibited when both are requested or Mode=1; automatic uses forward motion states only (PUB001, PUB002).
- Automatic motion: enabled by feed/cleaning/weighing/firing completion and held until the destination sensor is active; same-scan arrival has priority over completion (PUB003-PUB008).
- kick: set when weighing completes with weight<100.0 or weight>200.0; held while rejected until SensorWeight clears or Mode=0 (PUB009).
- firingTemp: updated only on a qualified weighing, REAL degrees, linear 100..200 -> 500..550; retained until an unqualified weighing or Mode=0 (PUB009, PUB010).
- CompletionLight: active while SensorOutput in automatic output state; cleared when the product is removed or Mode=0 (PUB008).
- Weight boundary test is inclusive: qualified is 100.0 <= weight <= 200.0 (PUB009).
*)
(* CONTRACT_RULES [] *)

TYPE E_ProductionState :
(
    ST_IDLE := 0,
    ST_MOVE_TO_WASH := 1,
    ST_AT_WASH := 2,
    ST_MOVE_TO_WEIGHT := 3,
    ST_AT_WEIGHT := 4,
    ST_MOVE_TO_FIRING := 5,
    ST_AT_FIRING := 6,
    ST_MOVE_TO_OUTPUT := 7,
    ST_AT_OUTPUT := 8,
    ST_REJECTED := 9
);
END_TYPE;

FUNCTION_BLOCK ProductionControl
VAR_INPUT
    Mode : BOOL;
    ForwardButton : BOOL;
    ReverseButton : BOOL;
    SensorFeed : BOOL;
    SensorWash : BOOL;
    SensorWeight : BOOL;
    SensorFiring : BOOL;
    SensorOutput : BOOL;
    washComplete : BOOL;
    weightComplete : BOOL;
    weight : REAL;
    firingComplete : BOOL;
END_VAR
VAR_OUTPUT
    MotorForward : BOOL;
    MotorReverse : BOOL;
    kick : BOOL;
    CompletionLight : BOOL;
    firingTemp : REAL;
END_VAR
VAR
    tmp_LocalState : E_ProductionState := ST_IDLE;
    tmp_Qualified : BOOL;
    tmp_TempLatched : REAL := 0.0;
END_VAR

IF NOT Mode THEN
    MotorForward := ForwardButton AND NOT ReverseButton;
    MotorReverse := ReverseButton AND NOT ForwardButton;
    kick := FALSE;
    CompletionLight := FALSE;
    tmp_TempLatched := 0.0;
    firingTemp := 0.0;
ELSE
    MotorReverse := FALSE;

    IF tmp_LocalState = ST_IDLE THEN
        IF SensorFeed THEN
            tmp_LocalState := ST_MOVE_TO_WASH;
        END_IF;
    ELSIF tmp_LocalState = ST_MOVE_TO_WASH THEN
        IF SensorWash THEN
            tmp_LocalState := ST_AT_WASH;
        END_IF;
    ELSIF tmp_LocalState = ST_AT_WASH THEN
        IF SensorWeight THEN
            tmp_LocalState := ST_AT_WEIGHT;
        ELSIF washComplete THEN
            tmp_LocalState := ST_MOVE_TO_WEIGHT;
        END_IF;
    ELSIF tmp_LocalState = ST_MOVE_TO_WEIGHT THEN
        IF SensorWeight THEN
            tmp_LocalState := ST_AT_WEIGHT;
        END_IF;
    ELSIF tmp_LocalState = ST_AT_WEIGHT THEN
        IF SensorFiring THEN
            tmp_LocalState := ST_AT_FIRING;
        ELSIF weightComplete THEN
            tmp_Qualified := (weight >= 100.0) AND (weight <= 200.0);
            IF tmp_Qualified THEN
                tmp_TempLatched := 500.0 + ((weight - 100.0) * 50.0) / 100.0;
                tmp_LocalState := ST_MOVE_TO_FIRING;
            ELSE
                tmp_TempLatched := 0.0;
                tmp_LocalState := ST_REJECTED;
            END_IF;
        END_IF;
    ELSIF tmp_LocalState = ST_REJECTED THEN
        IF NOT SensorWeight THEN
            tmp_TempLatched := 0.0;
            tmp_LocalState := ST_IDLE;
        END_IF;
    ELSIF tmp_LocalState = ST_MOVE_TO_FIRING THEN
        IF SensorFiring THEN
            tmp_LocalState := ST_AT_FIRING;
        END_IF;
    ELSIF tmp_LocalState = ST_AT_FIRING THEN
        IF SensorOutput THEN
            tmp_LocalState := ST_AT_OUTPUT;
        ELSIF firingComplete THEN
            tmp_LocalState := ST_MOVE_TO_OUTPUT;
        END_IF;
    ELSIF tmp_LocalState = ST_MOVE_TO_OUTPUT THEN
        IF SensorOutput THEN
            tmp_LocalState := ST_AT_OUTPUT;
        END_IF;
    ELSIF tmp_LocalState = ST_AT_OUTPUT THEN
        IF NOT SensorOutput THEN
            tmp_LocalState := ST_IDLE;
        END_IF;
    END_IF;

    CASE tmp_LocalState OF
        ST_MOVE_TO_WASH,
        ST_MOVE_TO_WEIGHT,
        ST_MOVE_TO_FIRING,
        ST_MOVE_TO_OUTPUT:
            MotorForward := TRUE;
    ELSE
            MotorForward := FALSE;
    END_CASE;

    kick := (tmp_LocalState = ST_REJECTED);
    CompletionLight := (tmp_LocalState = ST_AT_OUTPUT) AND SensorOutput;
    firingTemp := tmp_TempLatched;
END_IF;
END_FUNCTION_BLOCK

(* ---- public-hard-06.candidate_04.st ---- *)
(* ENGINEERING_CONTRACT
- MotorForward/MotorReverse: manual direct from buttons, both inhibited when both are requested or Mode=1; automatic uses forward motion states only (PUB001, PUB002).
- Automatic motion: enabled by feed/cleaning/weighing/firing completion and held until the destination sensor is active; same-scan arrival has priority over completion (PUB003-PUB008).
- kick: set when weighing completes with weight<100.0 or weight>200.0; held while rejected until SensorWeight clears or Mode=0 (PUB009).
- firingTemp: updated only on a qualified weighing, REAL degrees, linear 100..200 -> 500..550; retained until Mode=0 (PUB009, PUB010).
- CompletionLight: active while SensorOutput in automatic output state; cleared when the product is removed or Mode=0 (PUB008).
- Weight boundary test is inclusive: qualified is 100.0 <= weight <= 200.0 (PUB009).
*)
(* CONTRACT_RULES [] *)

TYPE E_ProductionState :
(
    ST_IDLE := 0,
    ST_MOVE_TO_WASH := 1,
    ST_AT_WASH := 2,
    ST_MOVE_TO_WEIGHT := 3,
    ST_AT_WEIGHT := 4,
    ST_MOVE_TO_FIRING := 5,
    ST_AT_FIRING := 6,
    ST_MOVE_TO_OUTPUT := 7,
    ST_AT_OUTPUT := 8,
    ST_REJECTED := 9
);
END_TYPE;

FUNCTION_BLOCK ProductionControl
VAR_INPUT
    Mode : BOOL;
    ForwardButton : BOOL;
    ReverseButton : BOOL;
    SensorFeed : BOOL;
    SensorWash : BOOL;
    SensorWeight : BOOL;
    SensorFiring : BOOL;
    SensorOutput : BOOL;
    washComplete : BOOL;
    weightComplete : BOOL;
    weight : REAL;
    firingComplete : BOOL;
END_VAR
VAR_OUTPUT
    MotorForward : BOOL;
    MotorReverse : BOOL;
    kick : BOOL;
    CompletionLight : BOOL;
    firingTemp : REAL;
END_VAR
VAR
    tmp_LocalState : E_ProductionState := ST_IDLE;
    tmp_Qualified : BOOL;
    tmp_TempLatched : REAL := 0.0;
END_VAR

IF NOT Mode THEN
    MotorForward := ForwardButton AND NOT ReverseButton;
    MotorReverse := ReverseButton AND NOT ForwardButton;
    kick := FALSE;
    CompletionLight := FALSE;
    tmp_TempLatched := 0.0;
    firingTemp := 0.0;
ELSE
    MotorReverse := FALSE;

    IF tmp_LocalState = ST_IDLE THEN
        IF SensorFeed THEN
            tmp_LocalState := ST_MOVE_TO_WASH;
        END_IF;
    ELSIF tmp_LocalState = ST_MOVE_TO_WASH THEN
        IF SensorWash THEN
            tmp_LocalState := ST_AT_WASH;
        END_IF;
    ELSIF tmp_LocalState = ST_AT_WASH THEN
        IF SensorWeight THEN
            tmp_LocalState := ST_AT_WEIGHT;
        ELSIF washComplete THEN
            tmp_LocalState := ST_MOVE_TO_WEIGHT;
        END_IF;
    ELSIF tmp_LocalState = ST_MOVE_TO_WEIGHT THEN
        IF SensorWeight THEN
            tmp_LocalState := ST_AT_WEIGHT;
        END_IF;
    ELSIF tmp_LocalState = ST_AT_WEIGHT THEN
        IF SensorFiring THEN
            tmp_LocalState := ST_AT_FIRING;
        ELSIF weightComplete THEN
            tmp_Qualified := (weight >= 100.0) AND (weight <= 200.0);
            IF tmp_Qualified THEN
                tmp_TempLatched := 500.0 + ((weight - 100.0) * 50.0) / 100.0;
                tmp_LocalState := ST_MOVE_TO_FIRING;
            ELSE
                tmp_LocalState := ST_REJECTED;
            END_IF;
        END_IF;
    ELSIF tmp_LocalState = ST_REJECTED THEN
        IF NOT SensorWeight THEN
            tmp_TempLatched := 0.0;
            tmp_LocalState := ST_IDLE;
        END_IF;
    ELSIF tmp_LocalState = ST_MOVE_TO_FIRING THEN
        IF SensorFiring THEN
            tmp_LocalState := ST_AT_FIRING;
        END_IF;
    ELSIF tmp_LocalState = ST_AT_FIRING THEN
        IF SensorOutput THEN
            tmp_LocalState := ST_AT_OUTPUT;
        ELSIF firingComplete THEN
            tmp_LocalState := ST_MOVE_TO_OUTPUT;
        END_IF;
    ELSIF tmp_LocalState = ST_MOVE_TO_OUTPUT THEN
        IF SensorOutput THEN
            tmp_LocalState := ST_AT_OUTPUT;
        END_IF;
    ELSIF tmp_LocalState = ST_AT_OUTPUT THEN
        IF NOT SensorOutput THEN
            tmp_LocalState := ST_IDLE;
        END_IF;
    END_IF;

    CASE tmp_LocalState OF
        ST_MOVE_TO_WASH,
        ST_MOVE_TO_WEIGHT,
        ST_MOVE_TO_FIRING,
        ST_MOVE_TO_OUTPUT:
            MotorForward := TRUE;
    ELSE
            MotorForward := FALSE;
    END_CASE;

    kick := (tmp_LocalState = ST_REJECTED);
    CompletionLight := (tmp_LocalState = ST_AT_OUTPUT) AND SensorOutput;
    firingTemp := tmp_TempLatched;
END_IF;
END_FUNCTION_BLOCK

(* ---- public-hard-06.patch_base_02.st ---- *)
(* ENGINEERING_CONTRACT
- MotorForward/MotorReverse: manual direct from buttons, both inhibited when both are requested or Mode=1; automatic uses forward motion states only (PUB001, PUB002).
- Automatic motion: enabled by feed/cleaning/weighing/firing completion and held until the destination sensor is active; same-scan arrival has priority over completion (PUB003-PUB008).
- kick: set when weighing completes with weight<100.0 or weight>200.0; held while rejected until SensorWeight clears or Mode=0 (PUB009).
- firingTemp: updated only on a qualified weighing, REAL degrees, linear 100..200 -> 500..550; held through firing/output until unqualified, next feed, or Mode=0 (PUB009, PUB010).
- CompletionLight: active while SensorOutput in automatic output state; cleared when the product is removed or Mode=0 (PUB008).
- Weight boundary test is inclusive: qualified is 100.0 <= weight <= 200.0 (PUB009).
*)
(* CONTRACT_RULES [] *)

TYPE E_ProductionState :
(
    ST_IDLE := 0,
    ST_MOVE_TO_WASH := 1,
    ST_AT_WASH := 2,
    ST_MOVE_TO_WEIGHT := 3,
    ST_AT_WEIGHT := 4,
    ST_MOVE_TO_FIRING := 5,
    ST_AT_FIRING := 6,
    ST_MOVE_TO_OUTPUT := 7,
    ST_AT_OUTPUT := 8,
    ST_REJECTED := 9
);
END_TYPE;

FUNCTION_BLOCK ProductionControl
VAR_INPUT
    Mode : BOOL;
    ForwardButton : BOOL;
    ReverseButton : BOOL;
    SensorFeed : BOOL;
    SensorWash : BOOL;
    SensorWeight : BOOL;
    SensorFiring : BOOL;
    SensorOutput : BOOL;
    washComplete : BOOL;
    weightComplete : BOOL;
    weight : REAL;
    firingComplete : BOOL;
END_VAR
VAR_OUTPUT
    MotorForward : BOOL;
    MotorReverse : BOOL;
    kick : BOOL;
    CompletionLight : BOOL;
    firingTemp : REAL;
END_VAR
VAR
    tmp_LocalState : E_ProductionState := ST_IDLE;
    tmp_Qualified : BOOL;
    tmp_TempLatched : REAL := 0.0;
END_VAR

IF NOT Mode THEN
    MotorForward := ForwardButton AND NOT ReverseButton;
    MotorReverse := ReverseButton AND NOT ForwardButton;
    kick := FALSE;
    CompletionLight := FALSE;
    tmp_TempLatched := 0.0;
    firingTemp := 0.0;
ELSE
    MotorReverse := FALSE;

    IF tmp_LocalState = ST_IDLE THEN
        tmp_TempLatched := 0.0;
        IF SensorFeed THEN
            tmp_LocalState := ST_MOVE_TO_WASH;
        END_IF;
    ELSIF tmp_LocalState = ST_MOVE_TO_WASH THEN
        IF SensorWash THEN
            tmp_LocalState := ST_AT_WASH;
        END_IF;
    ELSIF tmp_LocalState = ST_AT_WASH THEN
        IF SensorWeight THEN
            tmp_LocalState := ST_AT_WEIGHT;
        ELSIF washComplete THEN
            tmp_LocalState := ST_MOVE_TO_WEIGHT;
        END_IF;
    ELSIF tmp_LocalState = ST_MOVE_TO_WEIGHT THEN
        IF SensorWeight THEN
            tmp_LocalState := ST_AT_WEIGHT;
        END_IF;
    ELSIF tmp_LocalState = ST_AT_WEIGHT THEN
        IF SensorFiring THEN
            tmp_LocalState := ST_AT_FIRING;
        ELSIF weightComplete THEN
            tmp_Qualified := (weight >= 100.0) AND (weight <= 200.0);
            IF tmp_Qualified THEN
                tmp_TempLatched := 500.0 + ((weight - 100.0) * 50.0) / 100.0;
                tmp_LocalState := ST_MOVE_TO_FIRING;
            ELSE
                tmp_TempLatched := 0.0;
                tmp_LocalState := ST_REJECTED;
            END_IF;
        END_IF;
    ELSIF tmp_LocalState = ST_REJECTED THEN
        IF NOT SensorWeight THEN
            tmp_TempLatched := 0.0;
            tmp_LocalState := ST_IDLE;
        END_IF;
    ELSIF tmp_LocalState = ST_MOVE_TO_FIRING THEN
        IF SensorFiring THEN
            tmp_LocalState := ST_AT_FIRING;
        END_IF;
    ELSIF tmp_LocalState = ST_AT_FIRING THEN
        IF SensorOutput THEN
            tmp_LocalState := ST_AT_OUTPUT;
        ELSIF firingComplete THEN
            tmp_LocalState := ST_MOVE_TO_OUTPUT;
        END_IF;
    ELSIF tmp_LocalState = ST_MOVE_TO_OUTPUT THEN
        IF SensorOutput THEN
            tmp_LocalState := ST_AT_OUTPUT;
        END_IF;
    ELSIF tmp_LocalState = ST_AT_OUTPUT THEN
        IF NOT SensorOutput THEN
            tmp_TempLatched := 0.0;
            tmp_LocalState := ST_IDLE;
        END_IF;
    END_IF;

    CASE tmp_LocalState OF
        ST_MOVE_TO_WASH,
        ST_MOVE_TO_WEIGHT,
        ST_MOVE_TO_FIRING,
        ST_MOVE_TO_OUTPUT:
            MotorForward := TRUE;
    ELSE
            MotorForward := FALSE;
    END_CASE;

    kick := (tmp_LocalState = ST_REJECTED);
    CompletionLight := (tmp_LocalState = ST_AT_OUTPUT) AND SensorOutput;
    firingTemp := tmp_TempLatched;
END_IF;

(* ---- public-hard-06.patch_base_03.st ---- *)
(* ENGINEERING_CONTRACT
- MotorForward/MotorReverse: manual direct from buttons, both inhibited when both are requested or Mode=1; automatic uses forward motion states only (PUB001, PUB002).
- Automatic motion: enabled by feed/cleaning/weighing/firing completion and held until the destination sensor is active; same-scan arrival has priority over completion (PUB003-PUB008).
- kick: set when weighing completes with weight<100.0 or weight>200.0; held while rejected until SensorWeight clears or Mode=0 (PUB009).
- firingTemp: updated only on a qualified weighing, REAL degrees, linear 100..200 -> 500..550; held through firing/output until unqualified, next feed, or Mode=0 (PUB009, PUB010).
- CompletionLight: active while SensorOutput in automatic output state; cleared when the product is removed or Mode=0 (PUB008).
- Weight boundary test is inclusive: qualified is 100.0 <= weight <= 200.0 (PUB009).
*)
(* CONTRACT_RULES [] *)

TYPE E_ProductionState :
(
    ST_IDLE := 0,
    ST_MOVE_TO_WASH := 1,
    ST_AT_WASH := 2,
    ST_MOVE_TO_WEIGHT := 3,
    ST_AT_WEIGHT := 4,
    ST_MOVE_TO_FIRING := 5,
    ST_AT_FIRING := 6,
    ST_MOVE_TO_OUTPUT := 7,
    ST_AT_OUTPUT := 8,
    ST_REJECTED := 9
);
END_TYPE;

FUNCTION_BLOCK ProductionControl
VAR_INPUT
    Mode : BOOL;
    ForwardButton : BOOL;
    ReverseButton : BOOL;
    SensorFeed : BOOL;
    SensorWash : BOOL;
    SensorWeight : BOOL;
    SensorFiring : BOOL;
    SensorOutput : BOOL;
    washComplete : BOOL;
    weightComplete : BOOL;
    weight : REAL;
    firingComplete : BOOL;
END_VAR
VAR_OUTPUT
    MotorForward : BOOL;
    MotorReverse : BOOL;
    kick : BOOL;
    CompletionLight : BOOL;
    firingTemp : REAL;
END_VAR
VAR
    tmp_LocalState : E_ProductionState := ST_IDLE;
    tmp_Qualified : BOOL;
    tmp_TempLatched : REAL := 0.0;
END_VAR

IF NOT Mode THEN
    MotorForward := ForwardButton AND NOT ReverseButton;
    MotorReverse := ReverseButton AND NOT ForwardButton;
    kick := FALSE;
    CompletionLight := FALSE;
    tmp_TempLatched := 0.0;
    firingTemp := 0.0;
ELSE
    MotorReverse := FALSE;

    IF tmp_LocalState = ST_IDLE THEN
        tmp_TempLatched := 0.0;
        IF SensorFeed THEN
            tmp_LocalState := ST_MOVE_TO_WASH;
        END_IF;
    ELSIF tmp_LocalState = ST_MOVE_TO_WASH THEN
        IF SensorWash THEN
            tmp_LocalState := ST_AT_WASH;
        END_IF;
    ELSIF tmp_LocalState = ST_AT_WASH THEN
        IF SensorWeight THEN
            tmp_LocalState := ST_AT_WEIGHT;
        ELSIF washComplete THEN
            tmp_LocalState := ST_MOVE_TO_WEIGHT;
        END_IF;
    ELSIF tmp_LocalState = ST_MOVE_TO_WEIGHT THEN
        IF SensorWeight THEN
            tmp_LocalState := ST_AT_WEIGHT;
        END_IF;
    ELSIF tmp_LocalState = ST_AT_WEIGHT THEN
        IF SensorFiring THEN
            tmp_LocalState := ST_AT_FIRING;
        ELSIF weightComplete THEN
            tmp_Qualified := (weight >= 100.0) AND (weight <= 200.0);
            IF tmp_Qualified THEN
                tmp_TempLatched := 500.0 + ((weight - 100.0) * 50.0) / 100.0;
                tmp_LocalState := ST_MOVE_TO_FIRING;
            ELSE
                tmp_TempLatched := 0.0;
                tmp_LocalState := ST_REJECTED;
            END_IF;
        END_IF;
    ELSIF tmp_LocalState = ST_REJECTED THEN
        IF NOT SensorWeight THEN
            tmp_TempLatched := 0.0;
            tmp_LocalState := ST_IDLE;
        END_IF;
    ELSIF tmp_LocalState = ST_MOVE_TO_FIRING THEN
        IF SensorFiring THEN
            tmp_LocalState := ST_AT_FIRING;
        END_IF;
    ELSIF tmp_LocalState = ST_AT_FIRING THEN
        IF SensorOutput THEN
            tmp_LocalState := ST_AT_OUTPUT;
        ELSIF firingComplete THEN
            tmp_LocalState := ST_MOVE_TO_OUTPUT;
        END_IF;
    ELSIF tmp_LocalState = ST_MOVE_TO_OUTPUT THEN
        IF SensorOutput THEN
            tmp_LocalState := ST_AT_OUTPUT;
        END_IF;
    ELSIF tmp_LocalState = ST_AT_OUTPUT THEN
        IF NOT SensorOutput THEN
            tmp_TempLatched := 0.0;
            tmp_LocalState := ST_IDLE;
        END_IF;
    END_IF;

    CASE tmp_LocalState OF
        ST_MOVE_TO_WASH,
        ST_MOVE_TO_WEIGHT,
        ST_MOVE_TO_FIRING,
        ST_MOVE_TO_OUTPUT:
            MotorForward := TRUE;
    ELSE
            MotorForward := FALSE;
    END_CASE;

    kick := (tmp_LocalState = ST_REJECTED);
    CompletionLight := (tmp_LocalState = ST_AT_OUTPUT) AND SensorOutput;
    firingTemp := tmp_TempLatched;
END_IF;
END_FUNCTION_BLOCK

(* ---- public-hard-06.patch_base_04.st ---- *)
(* ENGINEERING_CONTRACT
- MotorForward/MotorReverse: manual direct from buttons, both inhibited when both are requested or Mode=1; automatic uses forward motion states only (PUB001, PUB002).
- Automatic motion: enabled by feed/cleaning/weighing/firing completion and held until the destination sensor is active; same-scan arrival has priority over completion (PUB003-PUB008).
- kick: set when weighing completes with weight<100.0 or weight>200.0; held while rejected until SensorWeight clears or Mode=0 (PUB009).
- firingTemp: updated only on a qualified weighing, REAL degrees, linear 100..200 -> 500..550; retained until an unqualified weighing or Mode=0 (PUB009, PUB010).
- CompletionLight: active while SensorOutput in automatic output state; cleared when the product is removed or Mode=0 (PUB008).
- Weight boundary test is inclusive: qualified is 100.0 <= weight <= 200.0 (PUB009).
*)
(* CONTRACT_RULES [] *)

TYPE E_ProductionState :
(
    ST_IDLE := 0,
    ST_MOVE_TO_WASH := 1,
    ST_AT_WASH := 2,
    ST_MOVE_TO_WEIGHT := 3,
    ST_AT_WEIGHT := 4,
    ST_MOVE_TO_FIRING := 5,
    ST_AT_FIRING := 6,
    ST_MOVE_TO_OUTPUT := 7,
    ST_AT_OUTPUT := 8,
    ST_REJECTED := 9
);
END_TYPE;

FUNCTION_BLOCK ProductionControl
VAR_INPUT
    Mode : BOOL;
    ForwardButton : BOOL;
    ReverseButton : BOOL;
    SensorFeed : BOOL;
    SensorWash : BOOL;
    SensorWeight : BOOL;
    SensorFiring : BOOL;
    SensorOutput : BOOL;
    washComplete : BOOL;
    weightComplete : BOOL;
    weight : REAL;
    firingComplete : BOOL;
END_VAR
VAR_OUTPUT
    MotorForward : BOOL;
    MotorReverse : BOOL;
    kick : BOOL;
    CompletionLight : BOOL;
    firingTemp : REAL;
END_VAR
VAR
    tmp_LocalState : E_ProductionState := ST_IDLE;
    tmp_Qualified : BOOL;
    tmp_TempLatched : REAL := 0.0;
END_VAR

IF NOT Mode THEN
    MotorForward := ForwardButton AND NOT ReverseButton;
    MotorReverse := ReverseButton AND NOT ForwardButton;
    kick := FALSE;
    CompletionLight := FALSE;
    tmp_TempLatched := 0.0;
    firingTemp := 0.0;
ELSE
    MotorReverse := FALSE;

    IF tmp_LocalState = ST_IDLE THEN
        IF SensorFeed THEN
            tmp_LocalState := ST_MOVE_TO_WASH;
        END_IF;
    ELSIF tmp_LocalState = ST_MOVE_TO_WASH THEN
        IF SensorWash THEN
            tmp_LocalState := ST_AT_WASH;
        END_IF;
    ELSIF tmp_LocalState = ST_AT_WASH THEN
        IF SensorWeight THEN
            tmp_LocalState := ST_AT_WEIGHT;
        ELSIF washComplete THEN
            tmp_LocalState := ST_MOVE_TO_WEIGHT;
        END_IF;
    ELSIF tmp_LocalState = ST_MOVE_TO_WEIGHT THEN
        IF SensorWeight THEN
            tmp_LocalState := ST_AT_WEIGHT;
        END_IF;
    ELSIF tmp_LocalState = ST_AT_WEIGHT THEN
        IF SensorFiring THEN
            tmp_LocalState := ST_AT_FIRING;
        ELSIF weightComplete THEN
            tmp_Qualified := (weight >= 100.0) AND (weight <= 200.0);
            IF tmp_Qualified THEN
                tmp_TempLatched := 500.0 + ((weight - 100.0) * 50.0) / 100.0;
                tmp_LocalState := ST_MOVE_TO_FIRING;
            ELSE
                tmp_TempLatched := 0.0;
                tmp_LocalState := ST_REJECTED;
            END_IF;
        END_IF;
    ELSIF tmp_LocalState = ST_REJECTED THEN
        IF NOT SensorWeight THEN
            tmp_TempLatched := 0.0;
            tmp_LocalState := ST_IDLE;
        END_IF;
    ELSIF tmp_LocalState = ST_MOVE_TO_FIRING THEN
        IF SensorFiring THEN
            tmp_LocalState := ST_AT_FIRING;
        END_IF;
    ELSIF tmp_LocalState = ST_AT_FIRING THEN
        IF SensorOutput THEN
            tmp_LocalState := ST_AT_OUTPUT;
        ELSIF firingComplete THEN
            tmp_LocalState := ST_MOVE_TO_OUTPUT;
        END_IF;
    ELSIF tmp_LocalState = ST_MOVE_TO_OUTPUT THEN
        IF SensorOutput THEN
            tmp_LocalState := ST_AT_OUTPUT;
        END_IF;
    ELSIF tmp_LocalState = ST_AT_OUTPUT THEN
        IF NOT SensorOutput THEN
            tmp_LocalState := ST_IDLE;
        END_IF;
    END_IF;

    CASE tmp_LocalState OF
        ST_MOVE_TO_WASH,
        ST_MOVE_TO_WEIGHT,
        ST_MOVE_TO_FIRING,
        ST_MOVE_TO_OUTPUT:
            MotorForward := TRUE;
    ELSE
            MotorForward := FALSE;
    END_CASE;

    kick := (tmp_LocalState = ST_REJECTED);
    CompletionLight := (tmp_LocalState = ST_AT_OUTPUT) AND SensorOutput;
    firingTemp := tmp_TempLatched;
END_IF;
END_FUNCTION_BLOCK

(* ---- public-hard-06.raw_candidate_01.st ---- *)
(* ENGINEERING_CONTRACT
- MotorForward/MotorReverse: manual direct from buttons, both inhibited when both are requested or Mode=1; automatic uses forward motion states only (PUB001, PUB002).
- Automatic motion: enabled by feed/cleaning/weighing/firing completion and held until the destination sensor is active; same-scan arrival has priority over completion (PUB003-PUB008).
- kick: set when weighing completes with weight<100.0 or weight>200.0; held while rejected until SensorWeight clears or Mode=0 (PUB009).
- firingTemp: updated only on a qualified weighing, REAL degrees, linear 100..200 -> 500..550; held through firing/output until unqualified, next feed, or Mode=0 (PUB009, PUB010).
- CompletionLight: active while SensorOutput in automatic output state; cleared when the product is removed or Mode=0 (PUB008).
- Weight boundary test is inclusive: qualified is 100.0 <= weight <= 200.0 (PUB009).
*)
(* CONTRACT_RULES [] *)

TYPE E_ProductionState :
(
    ST_IDLE := 0,
    ST_MOVE_TO_WASH := 1,
    ST_AT_WASH := 2,
    ST_MOVE_TO_WEIGHT := 3,
    ST_AT_WEIGHT := 4,
    ST_MOVE_TO_FIRING := 5,
    ST_AT_FIRING := 6,
    ST_MOVE_TO_OUTPUT := 7,
    ST_AT_OUTPUT := 8,
    ST_REJECTED := 9
);
END_TYPE

FUNCTION_BLOCK ProductionControl
VAR_INPUT
    Mode : BOOL;
    ForwardButton : BOOL;
    ReverseButton : BOOL;
    SensorFeed : BOOL;
    SensorWash : BOOL;
    SensorWeight : BOOL;
    SensorFiring : BOOL;
    SensorOutput : BOOL;
    washComplete : BOOL;
    weightComplete : BOOL;
    weight : REAL;
    firingComplete : BOOL;
END_VAR
VAR_OUTPUT
    MotorForward : BOOL;
    MotorReverse : BOOL;
    kick : BOOL;
    CompletionLight : BOOL;
    firingTemp : REAL;
END_VAR
VAR
    tmp_LocalState : E_ProductionState := ST_IDLE;
    tmp_Qualified : BOOL;
    tmp_TempLatched : REAL := 0.0;
END_VAR

IF NOT Mode THEN
    MotorForward := ForwardButton AND NOT ReverseButton;
    MotorReverse := ReverseButton AND NOT ForwardButton;
    kick := FALSE;
    CompletionLight := FALSE;
    tmp_TempLatched := 0.0;
    firingTemp := 0.0;
ELSE
    MotorReverse := FALSE;

    IF tmp_LocalState = ST_IDLE THEN
        tmp_TempLatched := 0.0;
        IF SensorFeed THEN
            tmp_LocalState := ST_MOVE_TO_WASH;
        END_IF;
    ELSIF tmp_LocalState = ST_MOVE_TO_WASH THEN
        IF SensorWash THEN
            tmp_LocalState := ST_AT_WASH;
        END_IF;
    ELSIF tmp_LocalState = ST_AT_WASH THEN
        IF SensorWeight THEN
            tmp_LocalState := ST_AT_WEIGHT;
        ELSIF washComplete THEN
            tmp_LocalState := ST_MOVE_TO_WEIGHT;
        END_IF;
    ELSIF tmp_LocalState = ST_MOVE_TO_WEIGHT THEN
        IF SensorWeight THEN
            tmp_LocalState := ST_AT_WEIGHT;
        END_IF;
    ELSIF tmp_LocalState = ST_AT_WEIGHT THEN
        IF SensorFiring THEN
            tmp_LocalState := ST_AT_FIRING;
        ELSIF weightComplete THEN
            tmp_Qualified := (weight >= 100.0) AND (weight <= 200.0);
            IF tmp_Qualified THEN
                tmp_TempLatched := 500.0 + ((weight - 100.0) * 50.0) / 100.0;
                tmp_LocalState := ST_MOVE_TO_FIRING;
            ELSE
                tmp_TempLatched := 0.0;
                tmp_LocalState := ST_REJECTED;
            END_IF;
        END_IF;
    ELSIF tmp_LocalState = ST_REJECTED THEN
        IF NOT SensorWeight THEN
            tmp_TempLatched := 0.0;
            tmp_LocalState := ST_IDLE;
        END_IF;
    ELSIF tmp_LocalState = ST_MOVE_TO_FIRING THEN
        IF SensorFiring THEN
            tmp_LocalState := ST_AT_FIRING;
        END_IF;
    ELSIF tmp_LocalState = ST_AT_FIRING THEN
        IF SensorOutput THEN
            tmp_LocalState := ST_AT_OUTPUT;
        ELSIF firingComplete THEN
            tmp_LocalState := ST_MOVE_TO_OUTPUT;
        END_IF;
    ELSIF tmp_LocalState = ST_MOVE_TO_OUTPUT THEN
        IF SensorOutput THEN
            tmp_LocalState := ST_AT_OUTPUT;
        END_IF;
    ELSIF tmp_LocalState = ST_AT_OUTPUT THEN
        IF NOT SensorOutput THEN
            tmp_TempLatched := 0.0;
            tmp_LocalState := ST_IDLE;
        END_IF;
    END_IF;

    CASE tmp_LocalState OF
        ST_MOVE_TO_WASH,
        ST_MOVE_TO_WEIGHT,
        ST_MOVE_TO_FIRING,
        ST_MOVE_TO_OUTPUT:
            MotorForward := TRUE;
    ELSE
            MotorForward := FALSE;
    END_CASE;

    kick := (tmp_LocalState = ST_REJECTED);
    CompletionLight := (tmp_LocalState = ST_AT_OUTPUT) AND SensorOutput;
    firingTemp := tmp_TempLatched;
END_IF;

(* ---- public-hard-06.raw_candidate_02.st ---- *)
(* ENGINEERING_CONTRACT
- MotorForward/MotorReverse: manual direct from buttons, both inhibited when both are requested or Mode=1; automatic uses forward motion states only (PUB001, PUB002).
- Automatic motion: enabled by feed/cleaning/weighing/firing completion and held until the destination sensor is active; same-scan arrival has priority over completion (PUB003-PUB008).
- kick: set when weighing completes with weight<100.0 or weight>200.0; held while rejected until SensorWeight clears or Mode=0 (PUB009).
- firingTemp: updated only on a qualified weighing, REAL degrees, linear 100..200 -> 500..550; held through firing/output until unqualified, next feed, or Mode=0 (PUB009, PUB010).
- CompletionLight: active while SensorOutput in automatic output state; cleared when the product is removed or Mode=0 (PUB008).
- Weight boundary test is inclusive: qualified is 100.0 <= weight <= 200.0 (PUB009).
*)
(* CONTRACT_RULES [] *)

TYPE E_ProductionState :
(
    ST_IDLE := 0,
    ST_MOVE_TO_WASH := 1,
    ST_AT_WASH := 2,
    ST_MOVE_TO_WEIGHT := 3,
    ST_AT_WEIGHT := 4,
    ST_MOVE_TO_FIRING := 5,
    ST_AT_FIRING := 6,
    ST_MOVE_TO_OUTPUT := 7,
    ST_AT_OUTPUT := 8,
    ST_REJECTED := 9
);
END_TYPE;

FUNCTION_BLOCK ProductionControl
VAR_INPUT
    Mode : BOOL;
    ForwardButton : BOOL;
    ReverseButton : BOOL;
    SensorFeed : BOOL;
    SensorWash : BOOL;
    SensorWeight : BOOL;
    SensorFiring : BOOL;
    SensorOutput : BOOL;
    washComplete : BOOL;
    weightComplete : BOOL;
    weight : REAL;
    firingComplete : BOOL;
END_VAR
VAR_OUTPUT
    MotorForward : BOOL;
    MotorReverse : BOOL;
    kick : BOOL;
    CompletionLight : BOOL;
    firingTemp : REAL;
END_VAR
VAR
    tmp_LocalState : E_ProductionState := ST_IDLE;
    tmp_Qualified : BOOL;
    tmp_TempLatched : REAL := 0.0;
END_VAR

IF NOT Mode THEN
    MotorForward := ForwardButton AND NOT ReverseButton;
    MotorReverse := ReverseButton AND NOT ForwardButton;
    kick := FALSE;
    CompletionLight := FALSE;
    tmp_TempLatched := 0.0;
    firingTemp := 0.0;
ELSE
    MotorReverse := FALSE;

    IF tmp_LocalState = ST_IDLE THEN
        tmp_TempLatched := 0.0;
        IF SensorFeed THEN
            tmp_LocalState := ST_MOVE_TO_WASH;
        END_IF;
    ELSIF tmp_LocalState = ST_MOVE_TO_WASH THEN
        IF SensorWash THEN
            tmp_LocalState := ST_AT_WASH;
        END_IF;
    ELSIF tmp_LocalState = ST_AT_WASH THEN
        IF SensorWeight THEN
            tmp_LocalState := ST_AT_WEIGHT;
        ELSIF washComplete THEN
            tmp_LocalState := ST_MOVE_TO_WEIGHT;
        END_IF;
    ELSIF tmp_LocalState = ST_MOVE_TO_WEIGHT THEN
        IF SensorWeight THEN
            tmp_LocalState := ST_AT_WEIGHT;
        END_IF;
    ELSIF tmp_LocalState = ST_AT_WEIGHT THEN
        IF SensorFiring THEN
            tmp_LocalState := ST_AT_FIRING;
        ELSIF weightComplete THEN
            tmp_Qualified := (weight >= 100.0) AND (weight <= 200.0);
            IF tmp_Qualified THEN
                tmp_TempLatched := 500.0 + ((weight - 100.0) * 50.0) / 100.0;
                tmp_LocalState := ST_MOVE_TO_FIRING;
            ELSE
                tmp_TempLatched := 0.0;
                tmp_LocalState := ST_REJECTED;
            END_IF;
        END_IF;
    ELSIF tmp_LocalState = ST_REJECTED THEN
        IF NOT SensorWeight THEN
            tmp_TempLatched := 0.0;
            tmp_LocalState := ST_IDLE;
        END_IF;
    ELSIF tmp_LocalState = ST_MOVE_TO_FIRING THEN
        IF SensorFiring THEN
            tmp_LocalState := ST_AT_FIRING;
        END_IF;
    ELSIF tmp_LocalState = ST_AT_FIRING THEN
        IF SensorOutput THEN
            tmp_LocalState := ST_AT_OUTPUT;
        ELSIF firingComplete THEN
            tmp_LocalState := ST_MOVE_TO_OUTPUT;
        END_IF;
    ELSIF tmp_LocalState = ST_MOVE_TO_OUTPUT THEN
        IF SensorOutput THEN
            tmp_LocalState := ST_AT_OUTPUT;
        END_IF;
    ELSIF tmp_LocalState = ST_AT_OUTPUT THEN
        IF NOT SensorOutput THEN
            tmp_TempLatched := 0.0;
            tmp_LocalState := ST_IDLE;
        END_IF;
    END_IF;

    CASE tmp_LocalState OF
        ST_MOVE_TO_WASH,
        ST_MOVE_TO_WEIGHT,
        ST_MOVE_TO_FIRING,
        ST_MOVE_TO_OUTPUT:
            MotorForward := TRUE;
    ELSE
            MotorForward := FALSE;
    END_CASE;

    kick := (tmp_LocalState = ST_REJECTED);
    CompletionLight := (tmp_LocalState = ST_AT_OUTPUT) AND SensorOutput;
    firingTemp := tmp_TempLatched;
END_IF;
END_FUNCTION_BLOCK

(* ---- public-hard-06.raw_candidate_03.st ---- *)
(* ENGINEERING_CONTRACT
- MotorForward/MotorReverse: manual direct from buttons, both inhibited when both are requested or Mode=1; automatic uses forward motion states only (PUB001, PUB002).
- Automatic motion: enabled by feed/cleaning/weighing/firing completion and held until the destination sensor is active; same-scan arrival has priority over completion (PUB003-PUB008).
- kick: set when weighing completes with weight<100.0 or weight>200.0; held while rejected until SensorWeight clears or Mode=0 (PUB009).
- firingTemp: updated only on a qualified weighing, REAL degrees, linear 100..200 -> 500..550; retained until an unqualified weighing or Mode=0 (PUB009, PUB010).
- CompletionLight: active while SensorOutput in automatic output state; cleared when the product is removed or Mode=0 (PUB008).
- Weight boundary test is inclusive: qualified is 100.0 <= weight <= 200.0 (PUB009).
*)
(* CONTRACT_RULES [] *)

TYPE E_ProductionState :
(
    ST_IDLE := 0,
    ST_MOVE_TO_WASH := 1,
    ST_AT_WASH := 2,
    ST_MOVE_TO_WEIGHT := 3,
    ST_AT_WEIGHT := 4,
    ST_MOVE_TO_FIRING := 5,
    ST_AT_FIRING := 6,
    ST_MOVE_TO_OUTPUT := 7,
    ST_AT_OUTPUT := 8,
    ST_REJECTED := 9
);
END_TYPE;

FUNCTION_BLOCK ProductionControl
VAR_INPUT
    Mode : BOOL;
    ForwardButton : BOOL;
    ReverseButton : BOOL;
    SensorFeed : BOOL;
    SensorWash : BOOL;
    SensorWeight : BOOL;
    SensorFiring : BOOL;
    SensorOutput : BOOL;
    washComplete : BOOL;
    weightComplete : BOOL;
    weight : REAL;
    firingComplete : BOOL;
END_VAR
VAR_OUTPUT
    MotorForward : BOOL;
    MotorReverse : BOOL;
    kick : BOOL;
    CompletionLight : BOOL;
    firingTemp : REAL;
END_VAR
VAR
    tmp_LocalState : E_ProductionState := ST_IDLE;
    tmp_Qualified : BOOL;
    tmp_TempLatched : REAL := 0.0;
END_VAR

IF NOT Mode THEN
    MotorForward := ForwardButton AND NOT ReverseButton;
    MotorReverse := ReverseButton AND NOT ForwardButton;
    kick := FALSE;
    CompletionLight := FALSE;
    tmp_TempLatched := 0.0;
    firingTemp := 0.0;
ELSE
    MotorReverse := FALSE;

    IF tmp_LocalState = ST_IDLE THEN
        IF SensorFeed THEN
            tmp_LocalState := ST_MOVE_TO_WASH;
        END_IF;
    ELSIF tmp_LocalState = ST_MOVE_TO_WASH THEN
        IF SensorWash THEN
            tmp_LocalState := ST_AT_WASH;
        END_IF;
    ELSIF tmp_LocalState = ST_AT_WASH THEN
        IF SensorWeight THEN
            tmp_LocalState := ST_AT_WEIGHT;
        ELSIF washComplete THEN
            tmp_LocalState := ST_MOVE_TO_WEIGHT;
        END_IF;
    ELSIF tmp_LocalState = ST_MOVE_TO_WEIGHT THEN
        IF SensorWeight THEN
            tmp_LocalState := ST_AT_WEIGHT;
        END_IF;
    ELSIF tmp_LocalState = ST_AT_WEIGHT THEN
        IF SensorFiring THEN
            tmp_LocalState := ST_AT_FIRING;
        ELSIF weightComplete THEN
            tmp_Qualified := (weight >= 100.0) AND (weight <= 200.0);
            IF tmp_Qualified THEN
                tmp_TempLatched := 500.0 + ((weight - 100.0) * 50.0) / 100.0;
                tmp_LocalState := ST_MOVE_TO_FIRING;
            ELSE
                tmp_TempLatched := 0.0;
                tmp_LocalState := ST_REJECTED;
            END_IF;
        END_IF;
    ELSIF tmp_LocalState = ST_REJECTED THEN
        IF NOT SensorWeight THEN
            tmp_TempLatched := 0.0;
            tmp_LocalState := ST_IDLE;
        END_IF;
    ELSIF tmp_LocalState = ST_MOVE_TO_FIRING THEN
        IF SensorFiring THEN
            tmp_LocalState := ST_AT_FIRING;
        END_IF;
    ELSIF tmp_LocalState = ST_AT_FIRING THEN
        IF SensorOutput THEN
            tmp_LocalState := ST_AT_OUTPUT;
        ELSIF firingComplete THEN
            tmp_LocalState := ST_MOVE_TO_OUTPUT;
        END_IF;
    ELSIF tmp_LocalState = ST_MOVE_TO_OUTPUT THEN
        IF SensorOutput THEN
            tmp_LocalState := ST_AT_OUTPUT;
        END_IF;
    ELSIF tmp_LocalState = ST_AT_OUTPUT THEN
        IF NOT SensorOutput THEN
            tmp_LocalState := ST_IDLE;
        END_IF;
    END_IF;

    CASE tmp_LocalState OF
        ST_MOVE_TO_WASH,
        ST_MOVE_TO_WEIGHT,
        ST_MOVE_TO_FIRING,
        ST_MOVE_TO_OUTPUT:
            MotorForward := TRUE;
    ELSE
            MotorForward := FALSE;
    END_CASE;

    kick := (tmp_LocalState = ST_REJECTED);
    CompletionLight := (tmp_LocalState = ST_AT_OUTPUT) AND SensorOutput;
    firingTemp := tmp_TempLatched;
END_IF;
END_FUNCTION_BLOCK

(* ---- public-hard-06.raw_candidate_04.st ---- *)
(* ENGINEERING_CONTRACT
- MotorForward/MotorReverse: manual direct from buttons, both inhibited when both are requested or Mode=1; automatic uses forward motion states only (PUB001, PUB002).
- Automatic motion: enabled by feed/cleaning/weighing/firing completion and held until the destination sensor is active; same-scan arrival has priority over completion (PUB003-PUB008).
- kick: set when weighing completes with weight<100.0 or weight>200.0; held while rejected until SensorWeight clears or Mode=0 (PUB009).
- firingTemp: updated only on a qualified weighing, REAL degrees, linear 100..200 -> 500..550; retained until Mode=0 (PUB009, PUB010).
- CompletionLight: active while SensorOutput in automatic output state; cleared when the product is removed or Mode=0 (PUB008).
- Weight boundary test is inclusive: qualified is 100.0 <= weight <= 200.0 (PUB009).
*)
(* CONTRACT_RULES [] *)

TYPE E_ProductionState :
(
    ST_IDLE := 0,
    ST_MOVE_TO_WASH := 1,
    ST_AT_WASH := 2,
    ST_MOVE_TO_WEIGHT := 3,
    ST_AT_WEIGHT := 4,
    ST_MOVE_TO_FIRING := 5,
    ST_AT_FIRING := 6,
    ST_MOVE_TO_OUTPUT := 7,
    ST_AT_OUTPUT := 8,
    ST_REJECTED := 9
);
END_TYPE;

FUNCTION_BLOCK ProductionControl
VAR_INPUT
    Mode : BOOL;
    ForwardButton : BOOL;
    ReverseButton : BOOL;
    SensorFeed : BOOL;
    SensorWash : BOOL;
    SensorWeight : BOOL;
    SensorFiring : BOOL;
    SensorOutput : BOOL;
    washComplete : BOOL;
    weightComplete : BOOL;
    weight : REAL;
    firingComplete : BOOL;
END_VAR
VAR_OUTPUT
    MotorForward : BOOL;
    MotorReverse : BOOL;
    kick : BOOL;
    CompletionLight : BOOL;
    firingTemp : REAL;
END_VAR
VAR
    tmp_LocalState : E_ProductionState := ST_IDLE;
    tmp_Qualified : BOOL;
    tmp_TempLatched : REAL := 0.0;
END_VAR

IF NOT Mode THEN
    MotorForward := ForwardButton AND NOT ReverseButton;
    MotorReverse := ReverseButton AND NOT ForwardButton;
    kick := FALSE;
    CompletionLight := FALSE;
    tmp_TempLatched := 0.0;
    firingTemp := 0.0;
ELSE
    MotorReverse := FALSE;

    IF tmp_LocalState = ST_IDLE THEN
        IF SensorFeed THEN
            tmp_LocalState := ST_MOVE_TO_WASH;
        END_IF;
    ELSIF tmp_LocalState = ST_MOVE_TO_WASH THEN
        IF SensorWash THEN
            tmp_LocalState := ST_AT_WASH;
        END_IF;
    ELSIF tmp_LocalState = ST_AT_WASH THEN
        IF SensorWeight THEN
            tmp_LocalState := ST_AT_WEIGHT;
        ELSIF washComplete THEN
            tmp_LocalState := ST_MOVE_TO_WEIGHT;
        END_IF;
    ELSIF tmp_LocalState = ST_MOVE_TO_WEIGHT THEN
        IF SensorWeight THEN
            tmp_LocalState := ST_AT_WEIGHT;
        END_IF;
    ELSIF tmp_LocalState = ST_AT_WEIGHT THEN
        IF SensorFiring THEN
            tmp_LocalState := ST_AT_FIRING;
        ELSIF weightComplete THEN
            tmp_Qualified := (weight >= 100.0) AND (weight <= 200.0);
            IF tmp_Qualified THEN
                tmp_TempLatched := 500.0 + ((weight - 100.0) * 50.0) / 100.0;
                tmp_LocalState := ST_MOVE_TO_FIRING;
            ELSE
                tmp_LocalState := ST_REJECTED;
            END_IF;
        END_IF;
    ELSIF tmp_LocalState = ST_REJECTED THEN
        IF NOT SensorWeight THEN
            tmp_TempLatched := 0.0;
            tmp_LocalState := ST_IDLE;
        END_IF;
    ELSIF tmp_LocalState = ST_MOVE_TO_FIRING THEN
        IF SensorFiring THEN
            tmp_LocalState := ST_AT_FIRING;
        END_IF;
    ELSIF tmp_LocalState = ST_AT_FIRING THEN
        IF SensorOutput THEN
            tmp_LocalState := ST_AT_OUTPUT;
        ELSIF firingComplete THEN
            tmp_LocalState := ST_MOVE_TO_OUTPUT;
        END_IF;
    ELSIF tmp_LocalState = ST_MOVE_TO_OUTPUT THEN
        IF SensorOutput THEN
            tmp_LocalState := ST_AT_OUTPUT;
        END_IF;
    ELSIF tmp_LocalState = ST_AT_OUTPUT THEN
        IF NOT SensorOutput THEN
            tmp_LocalState := ST_IDLE;
        END_IF;
    END_IF;

    CASE tmp_LocalState OF
        ST_MOVE_TO_WASH,
        ST_MOVE_TO_WEIGHT,
        ST_MOVE_TO_FIRING,
        ST_MOVE_TO_OUTPUT:
            MotorForward := TRUE;
    ELSE
            MotorForward := FALSE;
    END_CASE;

    kick := (tmp_LocalState = ST_REJECTED);
    CompletionLight := (tmp_LocalState = ST_AT_OUTPUT) AND SensorOutput;
    firingTemp := tmp_TempLatched;
END_IF;
END_FUNCTION_BLOCK

(* ---- public-medium-01.candidate_01.st ---- *)
TYPE ST_Pump :
STRUCT
    priority : INT;
    selection : BOOL;
    RunComd : BOOL;
END_STRUCT
END_TYPE;

(* CONTRACT_RULES [] *)

FUNCTION_BLOCK FB_MultiPumpControl
VAR_INPUT
    mode : BOOL;
    start : BOOL;
    stop : BOOL;
END_VAR
VAR_IN_OUT
    pumpGroup : ARRAY[1..5] OF ST_Pump;
END_VAR
VAR
    RunEnabled : BOOL;
    tmp_i : INT;
    tmp_slot : INT;
    tmp_best : INT;
    tmp_best_priority : INT;
    tmp_found : BOOL;
    tmp_selected : ARRAY[1..5] OF BOOL;
END_VAR

(*
ENGINEERING_CONTRACT
RunComd[1..5]: active while RunEnabled and current operating-set membership is true; retained per scan only while that condition stays true; stop clears all commands; changing selection/top-3 set clears only no-longer-selected pumps; same-scan priority stop > start.
RunEnabled: activated by start; held until stop; explicit deactivation is stop only; stop has priority when start and stop are simultaneously asserted.
mode: FALSE = manual, command set is pumpGroup[i].selection; TRUE = automatic, command set is the 3 highest-priority pumps. Ties use lower array index 1..5.
Boundaries: fixed array 1..5; only RunComd is written.
PUB: PUB001-PUB004.
*)

IF stop THEN
    RunEnabled := FALSE;
ELSIF start THEN
    RunEnabled := TRUE;
END_IF;

IF mode THEN
    FOR tmp_i := 1 TO 5 DO
        tmp_selected[tmp_i] := FALSE;
    END_FOR;

    FOR tmp_slot := 1 TO 3 DO
        tmp_best := 0;
        tmp_best_priority := 0;
        tmp_found := FALSE;

        FOR tmp_i := 1 TO 5 DO
            IF NOT tmp_selected[tmp_i] THEN
                IF (NOT tmp_found) OR (pumpGroup[tmp_i].priority > tmp_best_priority) THEN
                    tmp_best := tmp_i;
                    tmp_best_priority := pumpGroup[tmp_i].priority;
                    tmp_found := TRUE;
                END_IF;
            END_IF;
        END_FOR;

        IF tmp_found THEN
            tmp_selected[tmp_best] := TRUE;
        END_IF;
    END_FOR;

    FOR tmp_i := 1 TO 5 DO
        pumpGroup[tmp_i].RunComd := tmp_selected[tmp_i] AND RunEnabled;
    END_FOR;
ELSE
    FOR tmp_i := 1 TO 5 DO
        pumpGroup[tmp_i].RunComd := pumpGroup[tmp_i].selection AND RunEnabled;
    END_FOR;
END_IF;

END_FUNCTION_BLOCK

(* ---- public-medium-01.raw_candidate_01.st ---- *)
TYPE ST_Pump :
STRUCT
    priority : INT;
    selection : BOOL;
    RunComd : BOOL;
END_STRUCT
END_TYPE

(* CONTRACT_RULES [] *)

FUNCTION_BLOCK FB_MultiPumpControl
VAR_INPUT
    mode : BOOL;
    start : BOOL;
    stop : BOOL;
END_VAR
VAR_IN_OUT
    pumpGroup : ARRAY[1..5] OF ST_Pump;
END_VAR
VAR
    RunEnabled : BOOL;
    tmp_i : INT;
    tmp_slot : INT;
    tmp_best : INT;
    tmp_best_priority : INT;
    tmp_found : BOOL;
    tmp_selected : ARRAY[1..5] OF BOOL;
END_VAR

(*
ENGINEERING_CONTRACT
RunComd[1..5]: active while RunEnabled and current operating-set membership is true; retained per scan only while that condition stays true; stop clears all commands; changing selection/top-3 set clears only no-longer-selected pumps; same-scan priority stop > start.
RunEnabled: activated by start; held until stop; explicit deactivation is stop only; stop has priority when start and stop are simultaneously asserted.
mode: FALSE = manual, command set is pumpGroup[i].selection; TRUE = automatic, command set is the 3 highest-priority pumps. Ties use lower array index 1..5.
Boundaries: fixed array 1..5; only RunComd is written.
PUB: PUB001-PUB004.
*)

IF stop THEN
    RunEnabled := FALSE;
ELSIF start THEN
    RunEnabled := TRUE;
END_IF;

IF mode THEN
    FOR tmp_i := 1 TO 5 DO
        tmp_selected[tmp_i] := FALSE;
    END_FOR;

    FOR tmp_slot := 1 TO 3 DO
        tmp_best := 0;
        tmp_best_priority := 0;
        tmp_found := FALSE;

        FOR tmp_i := 1 TO 5 DO
            IF NOT tmp_selected[tmp_i] THEN
                IF (NOT tmp_found) OR (pumpGroup[tmp_i].priority > tmp_best_priority) THEN
                    tmp_best := tmp_i;
                    tmp_best_priority := pumpGroup[tmp_i].priority;
                    tmp_found := TRUE;
                END_IF;
            END_IF;
        END_FOR;

        IF tmp_found THEN
            tmp_selected[tmp_best] := TRUE;
        END_IF;
    END_FOR;

    FOR tmp_i := 1 TO 5 DO
        pumpGroup[tmp_i].RunComd := tmp_selected[tmp_i] AND RunEnabled;
    END_FOR;
ELSE
    FOR tmp_i := 1 TO 5 DO
        pumpGroup[tmp_i].RunComd := pumpGroup[tmp_i].selection AND RunEnabled;
    END_FOR;
END_IF;

END_FUNCTION_BLOCK

(* ---- public-medium-02.candidate_01.st ---- *)
TYPE ST_AnalogChannel :
STRUCT
    enable : BOOL;
    hiLIM : REAL;
    loLIM : REAL;
    bipolar : BOOL;
    measuringMode : INT;
    retVal : WORD;
    outputValue : REAL;
END_STRUCT
END_TYPE;

FUNCTION_BLOCK AnalogBatchProcessing
VAR_INPUT
    count : DINT;
END_VAR
VAR_IN_OUT
    analogValues : ARRAY[*] OF INT;
    channels : ARRAY[*] OF ST_AnalogChannel;
END_VAR
VAR
    local_a_lower : DINT;
    local_a_upper : DINT;
    local_c_lower : DINT;
    local_c_upper : DINT;
    local_count : DINT;
    local_i : DINT;
    local_a_idx : DINT;
    local_c_idx : DINT;
    local_raw : INT;
    local_scaled : REAL;
END_VAR

(* ENGINEERING_CONTRACT
- Enabled channels convert; disabled channels retain prior retVal/outputValue (unspecified).
- Count selects the first count ordinal slots from each array lower bound; analog is read-only (PUB001, PUB002).
- Mode 0 maps unipolar raw 0..27648 or bipolar raw -27648..27648 linearly to loLIM..hiLIM; outside raw is extrapolated, not clamped (PUB003).
- Mode 1: outputValue = raw * 0.1. Mode 2: outputValue = raw * 0.01 (PUB004).
- Invalid mode sets 16#8001; hiLIM <= loLIM sets 16#8002. Mode error is checked first; error skips conversion/output update (PUB005, PUB006).
- Valid enabled conversion writes outputValue and retVal = 16#0000.
*)

(* CONTRACT_RULES [] *)

local_a_lower := LOWER_BOUND(analogValues, 1);
local_a_upper := UPPER_BOUND(analogValues, 1);
local_c_lower := LOWER_BOUND(channels, 1);
local_c_upper := UPPER_BOUND(channels, 1);

local_count := count;
IF local_count < 0 THEN
    local_count := 0;
END_IF;
IF local_count > (local_a_upper - local_a_lower + 1) THEN
    local_count := local_a_upper - local_a_lower + 1;
END_IF;
IF local_count > (local_c_upper - local_c_lower + 1) THEN
    local_count := local_c_upper - local_c_lower + 1;
END_IF;

FOR local_i := 0 TO local_count - 1 DO
    local_a_idx := local_a_lower + local_i;
    local_c_idx := local_c_lower + local_i;

    IF channels[local_c_idx].enable THEN
        IF channels[local_c_idx].measuringMode < 0
           OR channels[local_c_idx].measuringMode > 2 THEN
            channels[local_c_idx].retVal := 16#8001;
        ELSIF channels[local_c_idx].hiLIM <= channels[local_c_idx].loLIM THEN
            channels[local_c_idx].retVal := 16#8002;
        ELSE
            local_raw := analogValues[local_a_idx];

            CASE channels[local_c_idx].measuringMode OF
                0:
                    IF channels[local_c_idx].bipolar THEN
                        local_scaled := channels[local_c_idx].loLIM
                                        + ((TO_REAL(local_raw) + 27648.0) / 55296.0)
                                          * (channels[local_c_idx].hiLIM - channels[local_c_idx].loLIM);
                    ELSE
                        local_scaled := channels[local_c_idx].loLIM
                                        + (TO_REAL(local_raw) / 27648.0)
                                          * (channels[local_c_idx].hiLIM - channels[local_c_idx].loLIM);
                    END_IF;

                1:
                    local_scaled := TO_REAL(local_raw) * 0.1;

                2:
                    local_scaled := TO_REAL(local_raw) * 0.01;
            END_CASE;

            channels[local_c_idx].outputValue := local_scaled;
            channels[local_c_idx].retVal := 16#0000;
        END_IF;
    END_IF;
END_FOR;

END_FUNCTION_BLOCK

(* ---- public-medium-02.raw_candidate_01.st ---- *)
TYPE ST_AnalogChannel :
STRUCT
    enable : BOOL;
    hiLIM : REAL;
    loLIM : REAL;
    bipolar : BOOL;
    measuringMode : INT;
    retVal : WORD;
    outputValue : REAL;
END_STRUCT
END_TYPE

FUNCTION_BLOCK AnalogBatchProcessing
VAR_INPUT
    count : DINT;
END_VAR
VAR_IN_OUT
    analogValues : ARRAY[*] OF INT;
    channels : ARRAY[*] OF ST_AnalogChannel;
END_VAR
VAR
    local_a_lower : DINT;
    local_a_upper : DINT;
    local_c_lower : DINT;
    local_c_upper : DINT;
    local_count : DINT;
    local_i : DINT;
    local_a_idx : DINT;
    local_c_idx : DINT;
    local_raw : INT;
    local_scaled : REAL;
END_VAR

(* ENGINEERING_CONTRACT
- Enabled channels convert; disabled channels retain prior retVal/outputValue (unspecified).
- Count selects the first count ordinal slots from each array lower bound; analog is read-only (PUB001, PUB002).
- Mode 0 maps unipolar raw 0..27648 or bipolar raw -27648..27648 linearly to loLIM..hiLIM; outside raw is extrapolated, not clamped (PUB003).
- Mode 1: outputValue = raw * 0.1. Mode 2: outputValue = raw * 0.01 (PUB004).
- Invalid mode sets 16#8001; hiLIM <= loLIM sets 16#8002. Mode error is checked first; error skips conversion/output update (PUB005, PUB006).
- Valid enabled conversion writes outputValue and retVal = 16#0000.
*)

(* CONTRACT_RULES [] *)

local_a_lower := LOWER_BOUND(analogValues, 1);
local_a_upper := UPPER_BOUND(analogValues, 1);
local_c_lower := LOWER_BOUND(channels, 1);
local_c_upper := UPPER_BOUND(channels, 1);

local_count := count;
IF local_count < 0 THEN
    local_count := 0;
END_IF
IF local_count > (local_a_upper - local_a_lower + 1) THEN
    local_count := local_a_upper - local_a_lower + 1;
END_IF
IF local_count > (local_c_upper - local_c_lower + 1) THEN
    local_count := local_c_upper - local_c_lower + 1;
END_IF

FOR local_i := 0 TO local_count - 1 DO
    local_a_idx := local_a_lower + local_i;
    local_c_idx := local_c_lower + local_i;

    IF channels[local_c_idx].enable THEN
        IF channels[local_c_idx].measuringMode < 0
           OR channels[local_c_idx].measuringMode > 2 THEN
            channels[local_c_idx].retVal := 16#8001;
        ELSIF channels[local_c_idx].hiLIM <= channels[local_c_idx].loLIM THEN
            channels[local_c_idx].retVal := 16#8002;
        ELSE
            local_raw := analogValues[local_a_idx];

            CASE channels[local_c_idx].measuringMode OF
                0:
                    IF channels[local_c_idx].bipolar THEN
                        local_scaled := channels[local_c_idx].loLIM
                                        + ((TO_REAL(local_raw) + 27648.0) / 55296.0)
                                          * (channels[local_c_idx].hiLIM - channels[local_c_idx].loLIM);
                    ELSE
                        local_scaled := channels[local_c_idx].loLIM
                                        + (TO_REAL(local_raw) / 27648.0)
                                          * (channels[local_c_idx].hiLIM - channels[local_c_idx].loLIM);
                    END_IF

                1:
                    local_scaled := TO_REAL(local_raw) * 0.1;

                2:
                    local_scaled := TO_REAL(local_raw) * 0.01;
            END_CASE

            channels[local_c_idx].outputValue := local_scaled;
            channels[local_c_idx].retVal := 16#0000;
        END_IF
    END_IF
END_FOR

END_FUNCTION_BLOCK

(* ---- public-medium-03.candidate_01.st ---- *)
FUNCTION_BLOCK FB_MovingAverage
VAR_INPUT
    cyclicExecution : BOOL;
    trigger : BOOL;
    value : LREAL;
    windowSize : INT;
    reset : BOOL;
END_VAR
VAR_OUTPUT
    average : LREAL;
    windowSizeReached : BOOL;
    error : BOOL;
    status : WORD;
END_VAR
VAR
    local_buffer : ARRAY[0..99] OF LREAL;
    local_sampleCount : INT;
    local_nextWrite : INT;
    local_triggerPrevious : BOOL;
    local_windowValid : BOOL;
    local_update : BOOL;
    local_i : INT;
    local_age : INT;
    local_position : INT;
    local_sum : LREAL;
END_VAR

(* CONTRACT_RULES [] *)

(* ENGINEERING_CONTRACT
   average: updated after valid acquisition (PUB001/PUB002); recalculated while window valid; 0.0 on reset; retained on invalid/no-reset.
   windowSizeReached: TRUE when stored sample count >= windowSize; cleared by reset and invalid window (PUB006).
   error/status: combinational from 1..100 window check (PUB003/PUB004); 16#8200 wins over 16#0000.
   reset: level-active; clears history, average, reached; suppresses same-scan acquisition (PUB003).
   acquisition: cyclicExecution first (PUB001); trigger edge only when cyclicExecution is FALSE (PUB002).
   retention: last up to 100 samples retained; mean is over newest windowSize samples (PUB001/PUB006).
   boundaries: valid windowSize 1..100 inclusive; trigger edge consumed every scan to avoid stale queuing.
*)

local_windowValid := (windowSize >= 1) AND (windowSize <= 100);

IF local_windowValid THEN
    error := FALSE;
    status := 16#0000;
ELSE
    error := TRUE;
    status := 16#8200;
END_IF;

IF reset THEN
    local_sampleCount := 0;
    local_nextWrite := 0;
    average := 0.0;
    windowSizeReached := FALSE;

    FOR local_i := 0 TO 99 BY 1 DO
        local_buffer[local_i] := 0.0;
    END_FOR;
ELSE
    IF NOT local_windowValid THEN
        windowSizeReached := FALSE;
    ELSE
        local_update := FALSE;

        IF cyclicExecution THEN
            local_update := TRUE;
        ELSIF (trigger AND NOT local_triggerPrevious) THEN
            local_update := TRUE;
        END_IF;

        IF local_update THEN
            local_buffer[local_nextWrite] := value;
            local_nextWrite := (local_nextWrite + 1) MOD 100;

            IF local_sampleCount < 100 THEN
                local_sampleCount := local_sampleCount + 1;
            END_IF;
        END_IF;

        local_sum := 0.0;

        IF local_sampleCount >= windowSize THEN
            FOR local_i := 0 TO windowSize - 1 BY 1 DO
                local_age := windowSize - 1 - local_i;
                local_position := (local_nextWrite + 100 - 1 - local_age) MOD 100;
                local_sum := local_sum + local_buffer[local_position];
            END_FOR;

            average := local_sum / INT_TO_LREAL(windowSize);
            windowSizeReached := TRUE;
        ELSIF local_sampleCount > 0 THEN
            FOR local_i := 0 TO local_sampleCount - 1 BY 1 DO
                local_age := local_sampleCount - 1 - local_i;
                local_position := (local_nextWrite + 100 - 1 - local_age) MOD 100;
                local_sum := local_sum + local_buffer[local_position];
            END_FOR;

            average := local_sum / INT_TO_LREAL(local_sampleCount);
            windowSizeReached := FALSE;
        ELSE
            average := 0.0;
            windowSizeReached := FALSE;
        END_IF;
    END_IF;
END_IF;

local_triggerPrevious := trigger;

END_FUNCTION_BLOCK

(* ---- public-medium-03.raw_candidate_01.st ---- *)
FUNCTION_BLOCK FB_MovingAverage
VAR_INPUT
    cyclicExecution : BOOL;
    trigger : BOOL;
    value : LREAL;
    windowSize : INT;
    reset : BOOL;
END_VAR
VAR_OUTPUT
    average : LREAL;
    windowSizeReached : BOOL;
    error : BOOL;
    status : WORD;
END_VAR
VAR
    local_buffer : ARRAY[0..99] OF LREAL;
    local_sampleCount : INT;
    local_nextWrite : INT;
    local_triggerPrevious : BOOL;
    local_windowValid : BOOL;
    local_update : BOOL;
    local_i : INT;
    local_age : INT;
    local_position : INT;
    local_sum : LREAL;
END_VAR

(* CONTRACT_RULES [] *)

(* ENGINEERING_CONTRACT
   average: updated after valid acquisition (PUB001/PUB002); recalculated while window valid; 0.0 on reset; retained on invalid/no-reset.
   windowSizeReached: TRUE when stored sample count >= windowSize; cleared by reset and invalid window (PUB006).
   error/status: combinational from 1..100 window check (PUB003/PUB004); 16#8200 wins over 16#0000.
   reset: level-active; clears history, average, reached; suppresses same-scan acquisition (PUB003).
   acquisition: cyclicExecution first (PUB001); trigger edge only when cyclicExecution is FALSE (PUB002).
   retention: last up to 100 samples retained; mean is over newest windowSize samples (PUB001/PUB006).
   boundaries: valid windowSize 1..100 inclusive; trigger edge consumed every scan to avoid stale queuing.
*)

local_windowValid := (windowSize >= 1) AND (windowSize <= 100);

IF local_windowValid THEN
    error := FALSE;
    status := 16#0000;
ELSE
    error := TRUE;
    status := 16#8200;
END_IF;

IF reset THEN
    local_sampleCount := 0;
    local_nextWrite := 0;
    average := 0.0;
    windowSizeReached := FALSE;

    FOR local_i := 0 TO 99 BY 1 DO
        local_buffer[local_i] := 0.0;
    END_FOR;
ELSE
    IF NOT local_windowValid THEN
        windowSizeReached := FALSE;
    ELSE
        local_update := FALSE;

        IF cyclicExecution THEN
            local_update := TRUE;
        ELSIF (trigger AND NOT local_triggerPrevious) THEN
            local_update := TRUE;
        END_IF;

        IF local_update THEN
            local_buffer[local_nextWrite] := value;
            local_nextWrite := (local_nextWrite + 1) MOD 100;

            IF local_sampleCount < 100 THEN
                local_sampleCount := local_sampleCount + 1;
            END_IF;
        END_IF;

        local_sum := 0.0;

        IF local_sampleCount >= windowSize THEN
            FOR local_i := 0 TO windowSize - 1 BY 1 DO
                local_age := windowSize - 1 - local_i;
                local_position := (local_nextWrite + 100 - 1 - local_age) MOD 100;
                local_sum := local_sum + local_buffer[local_position];
            END_FOR;

            average := local_sum / INT_TO_LREAL(windowSize);
            windowSizeReached := TRUE;
        ELSIF local_sampleCount > 0 THEN
            FOR local_i := 0 TO local_sampleCount - 1 BY 1 DO
                local_age := local_sampleCount - 1 - local_i;
                local_position := (local_nextWrite + 100 - 1 - local_age) MOD 100;
                local_sum := local_sum + local_buffer[local_position];
            END_FOR;

            average := local_sum / INT_TO_LREAL(local_sampleCount);
            windowSizeReached := FALSE;
        ELSE
            average := 0.0;
            windowSizeReached := FALSE;
        END_IF;
    END_IF;
END_IF;

local_triggerPrevious := trigger;

END_FUNCTION_BLOCK

(* ---- public-medium-04.candidate_01.st ---- *)
FUNCTION_BLOCK FB
VAR_INPUT
    TemperatureSensorInput : REAL;
    SetTemperature : REAL;
END_VAR
VAR_OUTPUT
    CurrentTemperature : REAL;
    SetTempDisplay : REAL;
    HeaterStatus : BOOL;
    OverheatProtection : BOOL;
    HeaterOutput : BOOL;
END_VAR
VAR
    tmp_SensorFault : BOOL;
    tmp_HeaterRequest : BOOL;
    tmp_OverheatLatched : BOOL;
    tmp_WasOverheat : BOOL;
    tmp_ContinuityTimer : TON;
    tmp_CoolingTimer : TON;
END_VAR

(* ENGINEERING_CONTRACT
HeaterOutput:
  ACT: TemperatureSensorInput < SetTemperature, no sensor fault, no overheat [PUB003].
  HOLD: none; recalculated each scan. OFF: equal/higher setpoint, fault, or overheat [PUB004, PUB005, PUB007].
OverheatProtection:
  ACT: heater remains on continuously for >5s, latched; HOLD: latched; OFF: auto after T#3S cooldown [PUB005].
Displays:
  CurrentTemperature mirrors sensor, SetTempDisplay mirrors setpoint, HeaterStatus mirrors HeaterOutput,
  OverheatProtection mirrors overheat latch [PUB001, PUB006].
Priority same scan: fault and overheat inhibit HeaterOutput. Sensor fault: input <0.0 or >100.0.
Units: REAL temperature values, TIME 5s/3s. Equality/manual reset unspecified; equal setpoint turns heater off.
*)
(* CONTRACT_RULES [] *)

tmp_SensorFault := (TemperatureSensorInput < 0.0) OR (TemperatureSensorInput > 100.0);
CurrentTemperature := TemperatureSensorInput;
SetTempDisplay := SetTemperature;

tmp_WasOverheat := tmp_OverheatLatched;

IF tmp_WasOverheat THEN
    tmp_CoolingTimer(IN := TRUE, PT := T#3S);
    IF tmp_CoolingTimer.Q THEN
        tmp_OverheatLatched := FALSE;
    END_IF;
END_IF;

tmp_HeaterRequest := (NOT tmp_SensorFault) AND (NOT tmp_OverheatLatched) AND (TemperatureSensorInput < SetTemperature);
HeaterOutput := tmp_HeaterRequest;

tmp_ContinuityTimer(IN := HeaterOutput, PT := T#10S);
IF tmp_ContinuityTimer.ET > T#5S THEN
    tmp_OverheatLatched := TRUE;
    HeaterOutput := FALSE;
END_IF;

OverheatProtection := tmp_OverheatLatched;
HeaterStatus := HeaterOutput;

IF NOT tmp_WasOverheat THEN
    tmp_CoolingTimer(IN := tmp_OverheatLatched, PT := T#3S);
END_IF;
END_FUNCTION_BLOCK
